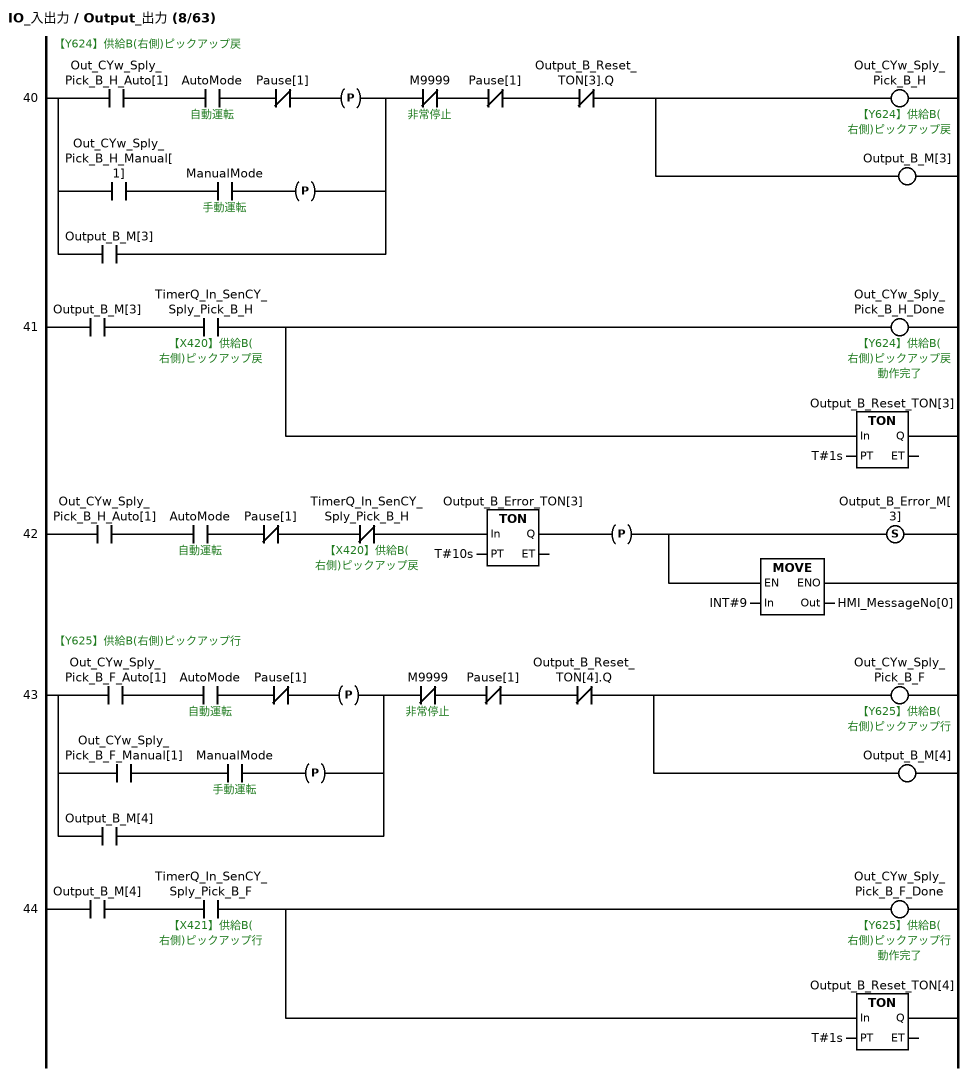
(* [picture p57: IO_入出力 / Output_出力, rungs 40-44] *)
(* Rung 40: 【Y624】供給B(右側)ピックアップ戻 *)
_e33(CLK := Out_CYw_Sply_Pick_B_H_Auto[1] AND AutoMode AND NOT Pause[1]);
_e34(CLK := Out_CYw_Sply_Pick_B_H_Manual[1] AND ManualMode);
_p35 := (_e33.Q OR _e34.Q OR Output_B_M[3]) AND NOT M9999 AND NOT Pause[1] AND NOT Output_B_Reset_TON[3].Q;
Out_CYw_Sply_Pick_B_H := _p35;
Output_B_M[3] := _p35;
(* Rung 41 *)
Out_CYw_Sply_Pick_B_H_Done := Output_B_M[3] AND TimerQ_In_SenCY_Sply_Pick_B_H;
Output_B_Reset_TON[3](In := Output_B_M[3] AND TimerQ_In_SenCY_Sply_Pick_B_H, PT := T#1s);
(* Rung 42 *)
Output_B_Error_TON[3](In := Out_CYw_Sply_Pick_B_H_Auto[1] AND AutoMode AND NOT Pause[1] AND NOT TimerQ_In_SenCY_Sply_Pick_B_H, PT := T#10s);
_e36(CLK := Output_B_Error_TON[3].Q);
IF _e36.Q THEN
    Output_B_Error_M[3] := TRUE;
    HMI_MessageNo[0] := INT#9;
END_IF;
(* Rung 43: 【Y625】供給B(右側)ピックアップ行 *)
_e37(CLK := Out_CYw_Sply_Pick_B_F_Auto[1] AND AutoMode AND NOT Pause[1]);
_e38(CLK := Out_CYw_Sply_Pick_B_F_Manual[1] AND ManualMode);
_p39 := (_e37.Q OR _e38.Q OR Output_B_M[4]) AND NOT M9999 AND NOT Pause[1] AND NOT Output_B_Reset_TON[4].Q;
Out_CYw_Sply_Pick_B_F := _p39;
Output_B_M[4] := _p39;
(* Rung 44 *)
Out_CYw_Sply_Pick_B_F_Done := Output_B_M[4] AND TimerQ_In_SenCY_Sply_Pick_B_F;
Output_B_Reset_TON[4](In := Output_B_M[4] AND TimerQ_In_SenCY_Sply_Pick_B_F, PT := T#1s);

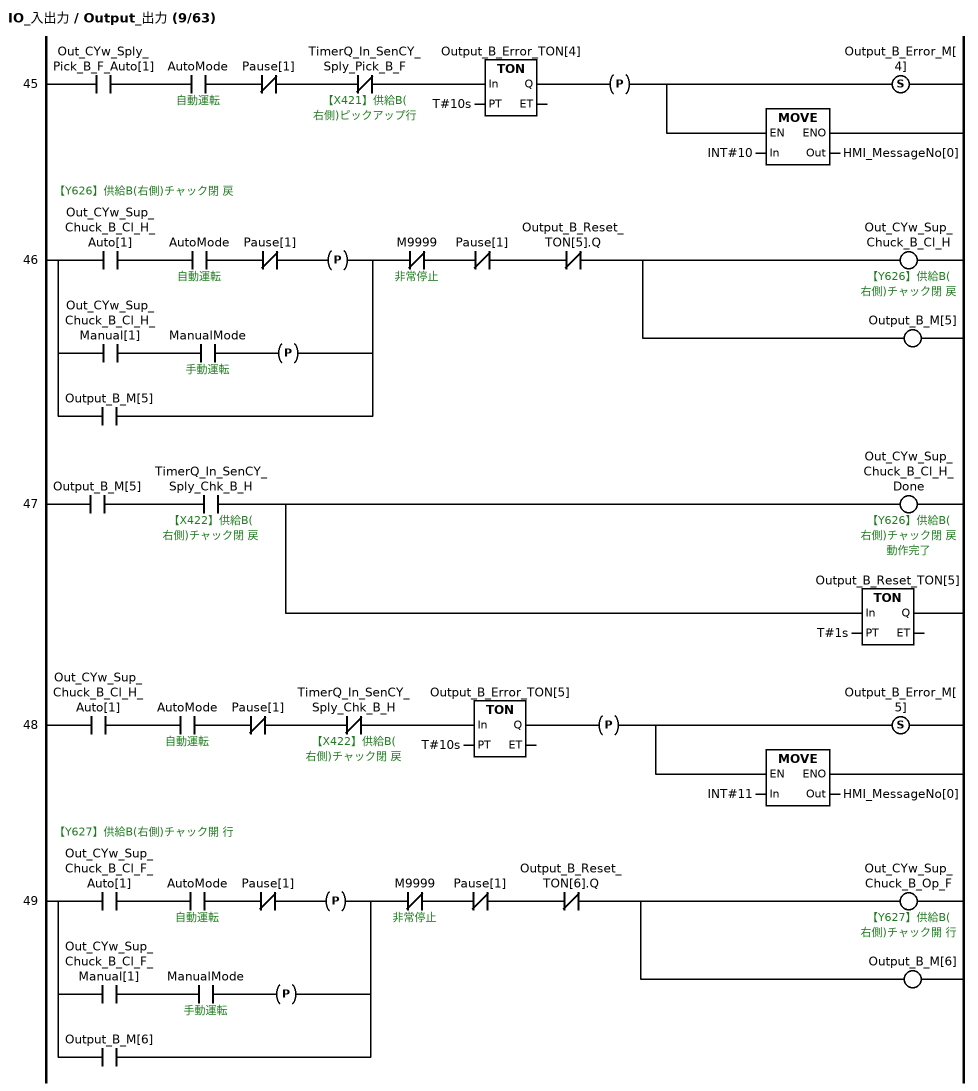
(* Rung 45 *)
Output_B_Error_TON[4](In := Out_CYw_Sply_Pick_B_F_Auto[1] AND AutoMode AND NOT Pause[1] AND NOT TimerQ_In_SenCY_Sply_Pick_B_F, PT := T#10s);
_e40(CLK := Output_B_Error_TON[4].Q);
IF _e40.Q THEN
    Output_B_Error_M[4] := TRUE;
    HMI_MessageNo[0] := INT#10;
END_IF;
(* Rung 46: 【Y626】供給B(右側)チャック閉 戻 *)
_e41(CLK := Out_CYw_Sup_Chuck_B_Cl_H_Auto[1] AND AutoMode AND NOT Pause[1]);
_e42(CLK := Out_CYw_Sup_Chuck_B_Cl_H_Manual[1] AND ManualMode);
_p43 := (_e41.Q OR _e42.Q OR Output_B_M[5]) AND NOT M9999 AND NOT Pause[1] AND NOT Output_B_Reset_TON[5].Q;
Out_CYw_Sup_Chuck_B_Cl_H := _p43;
Output_B_M[5] := _p43;
(* Rung 47 *)
Out_CYw_Sup_Chuck_B_Cl_H_Done := Output_B_M[5] AND TimerQ_In_SenCY_Sply_Chk_B_H;
Output_B_Reset_TON[5](In := Output_B_M[5] AND TimerQ_In_SenCY_Sply_Chk_B_H, PT := T#1s);
(* Rung 48 *)
Output_B_Error_TON[5](In := Out_CYw_Sup_Chuck_B_Cl_H_Auto[1] AND AutoMode AND NOT Pause[1] AND NOT TimerQ_In_SenCY_Sply_Chk_B_H, PT := T#10s);
_e44(CLK := Output_B_Error_TON[5].Q);
IF _e44.Q THEN
    Output_B_Error_M[5] := TRUE;
    HMI_MessageNo[0] := INT#11;
END_IF;
(* Rung 49: 【Y627】供給B(右側)チャック開 行 *)
_e45(CLK := Out_CYw_Sup_Chuck_B_Cl_F_Auto[1] AND AutoMode AND NOT Pause[1]);
_e46(CLK := Out_CYw_Sup_Chuck_B_Cl_F_Manual[1] AND ManualMode);
_p47 := (_e45.Q OR _e46.Q OR Output_B_M[6]) AND NOT M9999 AND NOT Pause[1] AND NOT Output_B_Reset_TON[6].Q;
Out_CYw_Sup_Chuck_B_Op_F := _p47;
Output_B_M[6] := _p47;

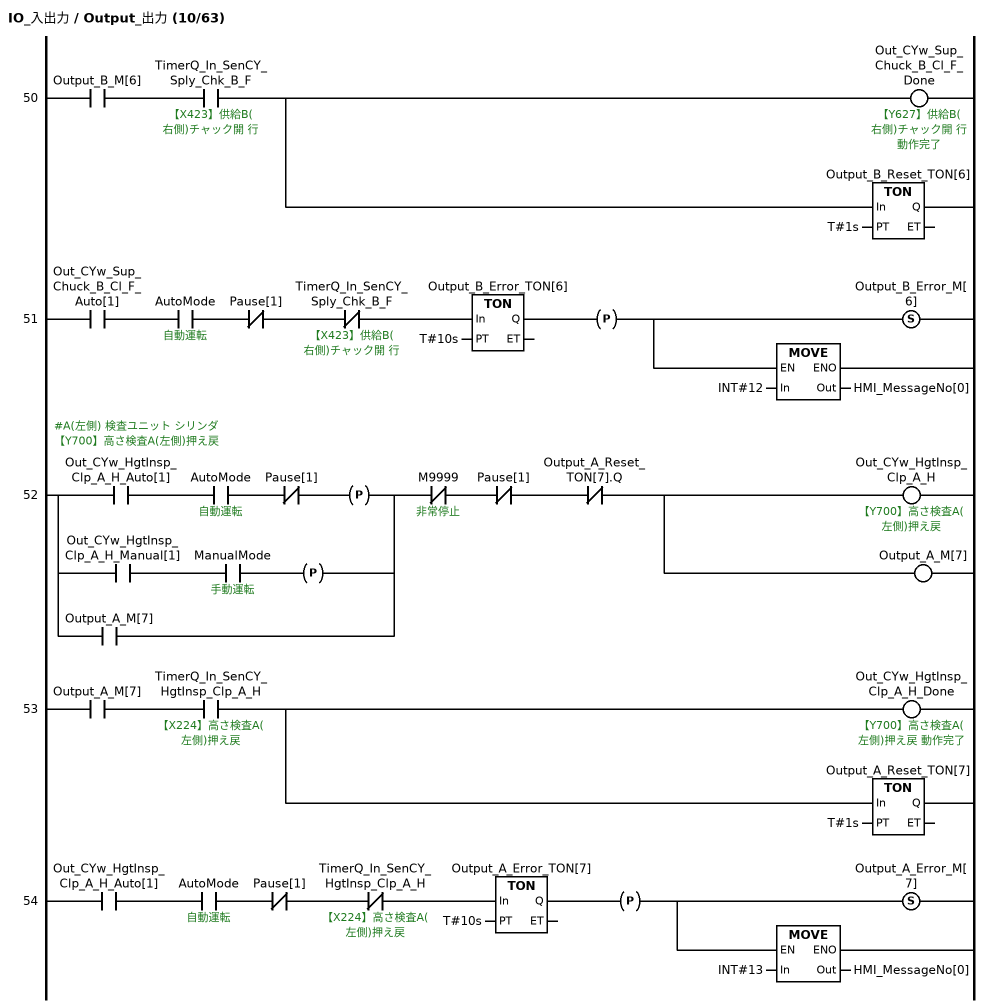
(* Rung 50 *)
Out_CYw_Sup_Chuck_B_Cl_F_Done := Output_B_M[6] AND TimerQ_In_SenCY_Sply_Chk_B_F;
Output_B_Reset_TON[6](In := Output_B_M[6] AND TimerQ_In_SenCY_Sply_Chk_B_F, PT := T#1s);
(* Rung 51 *)
Output_B_Error_TON[6](In := Out_CYw_Sup_Chuck_B_Cl_F_Auto[1] AND AutoMode AND NOT Pause[1] AND NOT TimerQ_In_SenCY_Sply_Chk_B_F, PT := T#10s);
_e48(CLK := Output_B_Error_TON[6].Q);
IF _e48.Q THEN
    Output_B_Error_M[6] := TRUE;
    HMI_MessageNo[0] := INT#12;
END_IF;
(* Rung 52: #A(左側) 検査ユニット シリンダ / 【Y700】高さ検査A(左側)押え戻 *)
_e49(CLK := Out_CYw_HgtInsp_Clp_A_H_Auto[1] AND AutoMode AND NOT Pause[1]);
_e50(CLK := Out_CYw_HgtInsp_Clp_A_H_Manual[1] AND ManualMode);
_p51 := (_e49.Q OR _e50.Q OR Output_A_M[7]) AND NOT M9999 AND NOT Pause[1] AND NOT Output_A_Reset_TON[7].Q;
Out_CYw_HgtInsp_Clp_A_H := _p51;
Output_A_M[7] := _p51;
(* Rung 53 *)
_p52 := Output_A_M[7] AND TimerQ_In_SenCY_HgtInsp_Clp_A_H;
Out_CYw_HgtInsp_Clp_A_H_Done := _p52;
Output_A_Reset_TON[7](In := _p52, PT := T#1s);
(* Rung 54 *)
Output_A_Error_TON[7](In := Out_CYw_HgtInsp_Clp_A_H_Auto[1] AND AutoMode AND NOT Pause[1] AND NOT TimerQ_In_SenCY_HgtInsp_Clp_A_H, PT := T#10s);
_e53(CLK := Output_A_Error_TON[7].Q);
IF _e53.Q THEN
    Output_A_Error_M[7] := TRUE;
    HMI_MessageNo[0] := INT#13;
END_IF;

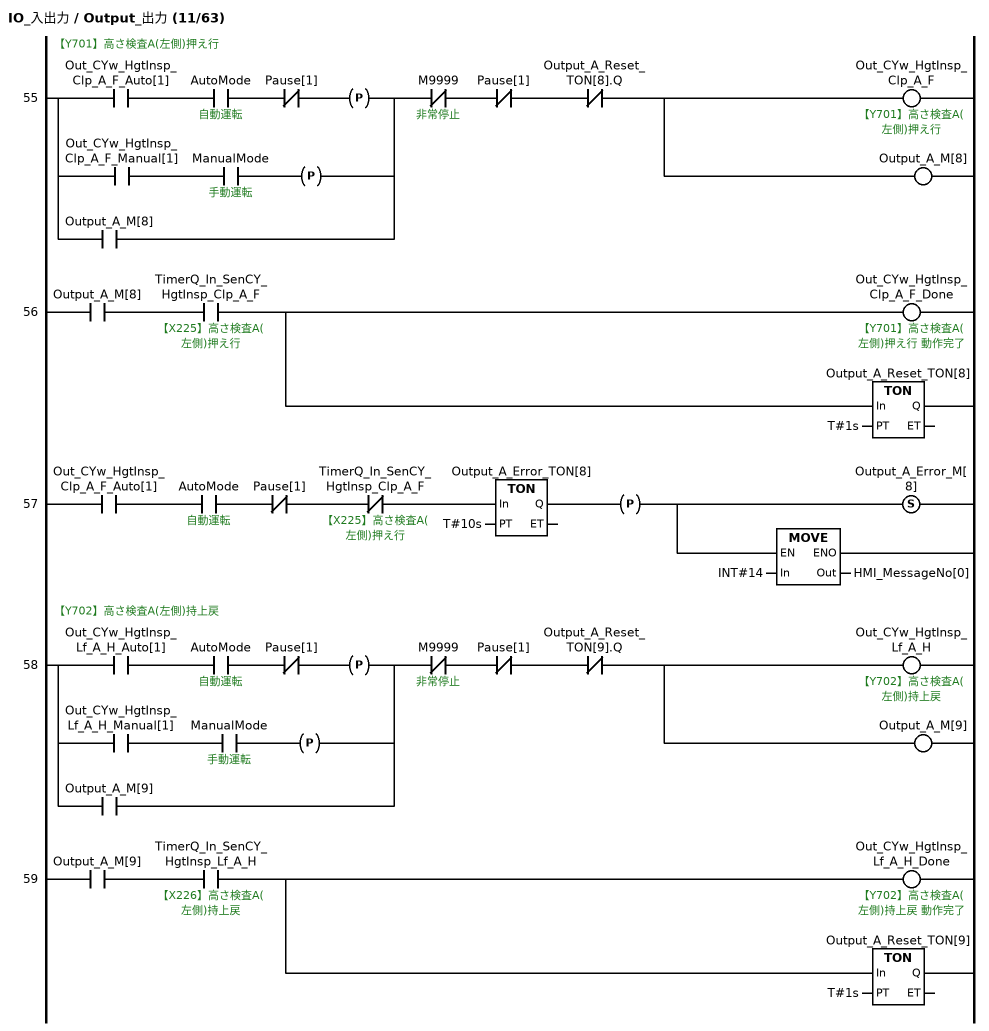
(* Rung 55: 【Y701】高さ検査A(左側)押え行 *)
_e54(CLK := Out_CYw_HgtInsp_Clp_A_F_Auto[1] AND AutoMode AND NOT Pause[1]);
_e55(CLK := Out_CYw_HgtInsp_Clp_A_F_Manual[1] AND ManualMode);
_p56 := (_e54.Q OR _e55.Q OR Output_A_M[8]) AND NOT M9999 AND NOT Pause[1] AND NOT Output_A_Reset_TON[8].Q;
Out_CYw_HgtInsp_Clp_A_F := _p56;
Output_A_M[8] := _p56;
(* Rung 56 *)
_p57 := Output_A_M[8] AND TimerQ_In_SenCY_HgtInsp_Clp_A_F;
Out_CYw_HgtInsp_Clp_A_F_Done := _p57;
Output_A_Reset_TON[8](In := _p57, PT := T#1s);
(* Rung 57 *)
Output_A_Error_TON[8](In := Out_CYw_HgtInsp_Clp_A_F_Auto[1] AND AutoMode AND NOT Pause[1] AND NOT TimerQ_In_SenCY_HgtInsp_Clp_A_F, PT := T#10s);
_e58(CLK := Output_A_Error_TON[8].Q);
IF _e58.Q THEN
    Output_A_Error_M[8] := TRUE;
    HMI_MessageNo[0] := INT#14;
END_IF;
(* Rung 58: 【Y702】高さ検査A(左側)持上戻 *)
_e59(CLK := Out_CYw_HgtInsp_Lf_A_H_Auto[1] AND AutoMode AND NOT Pause[1]);
_e60(CLK := Out_CYw_HgtInsp_Lf_A_H_Manual[1] AND ManualMode);
_p61 := (_e59.Q OR _e60.Q OR Output_A_M[9]) AND NOT M9999 AND NOT Pause[1] AND NOT Output_A_Reset_TON[9].Q;
Out_CYw_HgtInsp_Lf_A_H := _p61;
Output_A_M[9] := _p61;
(* Rung 59 *)
Out_CYw_HgtInsp_Lf_A_H_Done := Output_A_M[9] AND TimerQ_In_SenCY_HgtInsp_Lf_A_H;
Output_A_Reset_TON[9](In := Output_A_M[9] AND TimerQ_In_SenCY_HgtInsp_Lf_A_H, PT := T#1s);

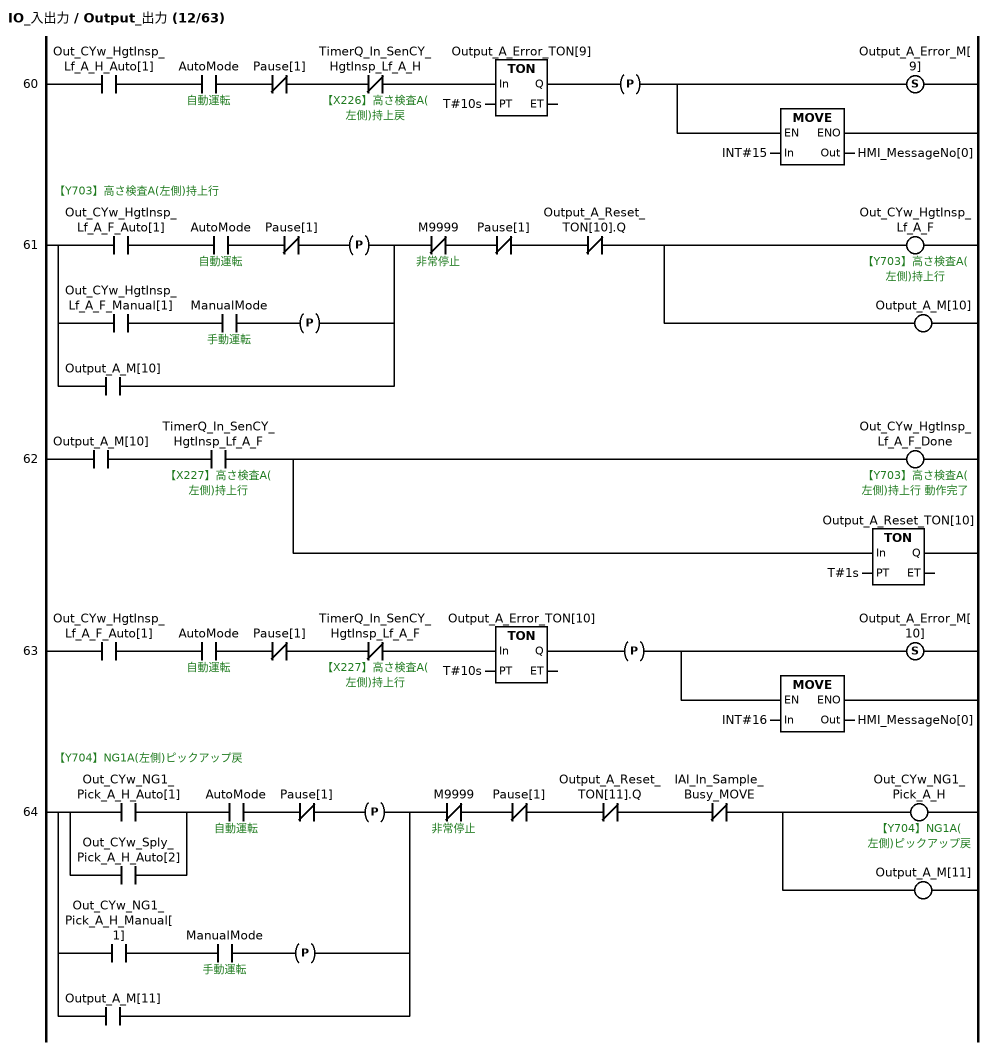
(* Rung 60 *)
Output_A_Error_TON[9](In := Out_CYw_HgtInsp_Lf_A_H_Auto[1] AND AutoMode AND NOT Pause[1] AND NOT TimerQ_In_SenCY_HgtInsp_Lf_A_H, PT := T#10s);
_e62(CLK := Output_A_Error_TON[9].Q);
IF _e62.Q THEN
    Output_A_Error_M[9] := TRUE;
    HMI_MessageNo[0] := INT#15;
END_IF;
(* Rung 61: 【Y703】高さ検査A(左側)持上行 *)
_e63(CLK := Out_CYw_HgtInsp_Lf_A_F_Auto[1] AND AutoMode AND NOT Pause[1]);
_e64(CLK := Out_CYw_HgtInsp_Lf_A_F_Manual[1] AND ManualMode);
_p65 := (_e63.Q OR _e64.Q OR Output_A_M[10]) AND NOT M9999 AND NOT Pause[1] AND NOT Output_A_Reset_TON[10].Q;
Out_CYw_HgtInsp_Lf_A_F := _p65;
Output_A_M[10] := _p65;
(* Rung 62 *)
_p66 := Output_A_M[10] AND TimerQ_In_SenCY_HgtInsp_Lf_A_F;
Out_CYw_HgtInsp_Lf_A_F_Done := _p66;
Output_A_Reset_TON[10](In := _p66, PT := T#1s);
(* Rung 63 *)
Output_A_Error_TON[10](In := Out_CYw_HgtInsp_Lf_A_F_Auto[1] AND AutoMode AND NOT Pause[1] AND NOT TimerQ_In_SenCY_HgtInsp_Lf_A_F, PT := T#10s);
_e67(CLK := Output_A_Error_TON[10].Q);
IF _e67.Q THEN
    Output_A_Error_M[10] := TRUE;
    HMI_MessageNo[0] := INT#16;
END_IF;
(* Rung 64: 【Y704】NG1A(左側)ピックアップ戻 *)
_e68(CLK := (Out_CYw_NG1_Pick_A_H_Auto[1] OR Out_CYw_Sply_Pick_A_H_Auto[2]) AND AutoMode AND NOT Pause[1]);
_e69(CLK := Out_CYw_NG1_Pick_A_H_Manual[1] AND ManualMode);
_p70 := (_e68.Q OR _e69.Q OR Output_A_M[11]) AND NOT M9999 AND NOT Pause[1] AND NOT Output_A_Reset_TON[11].Q AND NOT IAI_In_Sample_Busy_MOVE;
Out_CYw_NG1_Pick_A_H := _p70;
Output_A_M[11] := _p70;

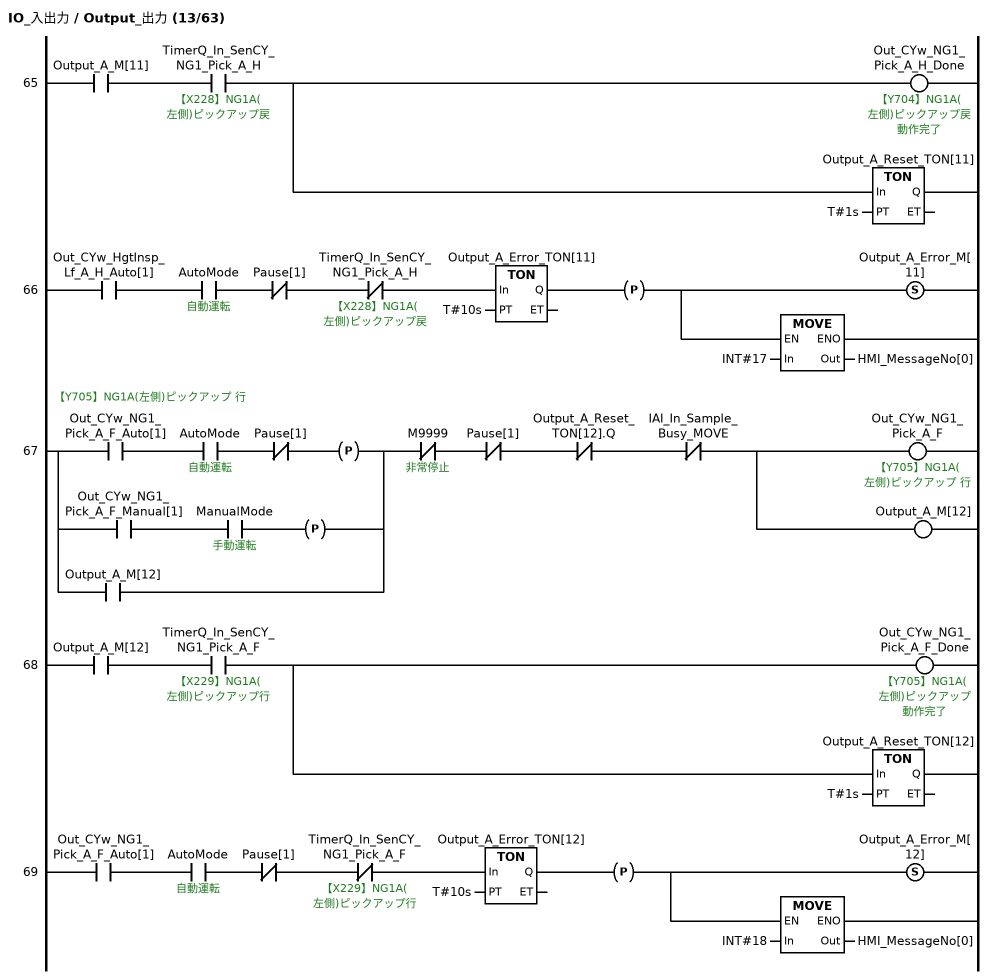
(* Rung 65 *)
Out_CYw_NG1_Pick_A_H_Done := Output_A_M[11] AND TimerQ_In_SenCY_NG1_Pick_A_H;
Output_A_Reset_TON[11](In := Output_A_M[11] AND TimerQ_In_SenCY_NG1_Pick_A_H, PT := T#1s);
(* Rung 66 *)
Output_A_Error_TON[11](In := Out_CYw_HgtInsp_Lf_A_H_Auto[1] AND AutoMode AND NOT Pause[1] AND NOT TimerQ_In_SenCY_NG1_Pick_A_H, PT := T#10s);
_e71(CLK := Output_A_Error_TON[11].Q);
IF _e71.Q THEN
    Output_A_Error_M[11] := TRUE;
    HMI_MessageNo[0] := INT#17;
END_IF;
(* Rung 67: 【Y705】NG1A(左側)ピックアップ 行 *)
_e72(CLK := Out_CYw_NG1_Pick_A_F_Auto[1] AND AutoMode AND NOT Pause[1]);
_e73(CLK := Out_CYw_NG1_Pick_A_F_Manual[1] AND ManualMode);
_p74 := (_e72.Q OR _e73.Q OR Output_A_M[12]) AND NOT M9999 AND NOT Pause[1] AND NOT Output_A_Reset_TON[12].Q AND NOT IAI_In_Sample_Busy_MOVE;
Out_CYw_NG1_Pick_A_F := _p74;
Output_A_M[12] := _p74;
(* Rung 68 *)
Out_CYw_NG1_Pick_A_F_Done := Output_A_M[12] AND TimerQ_In_SenCY_NG1_Pick_A_F;
Output_A_Reset_TON[12](In := Output_A_M[12] AND TimerQ_In_SenCY_NG1_Pick_A_F, PT := T#1s);
(* Rung 69 *)
Output_A_Error_TON[12](In := Out_CYw_NG1_Pick_A_F_Auto[1] AND AutoMode AND NOT Pause[1] AND NOT TimerQ_In_SenCY_NG1_Pick_A_F, PT := T#10s);
_e75(CLK := Output_A_Error_TON[12].Q);
IF _e75.Q THEN
    Output_A_Error_M[12] := TRUE;
    HMI_MessageNo[0] := INT#18;
END_IF;

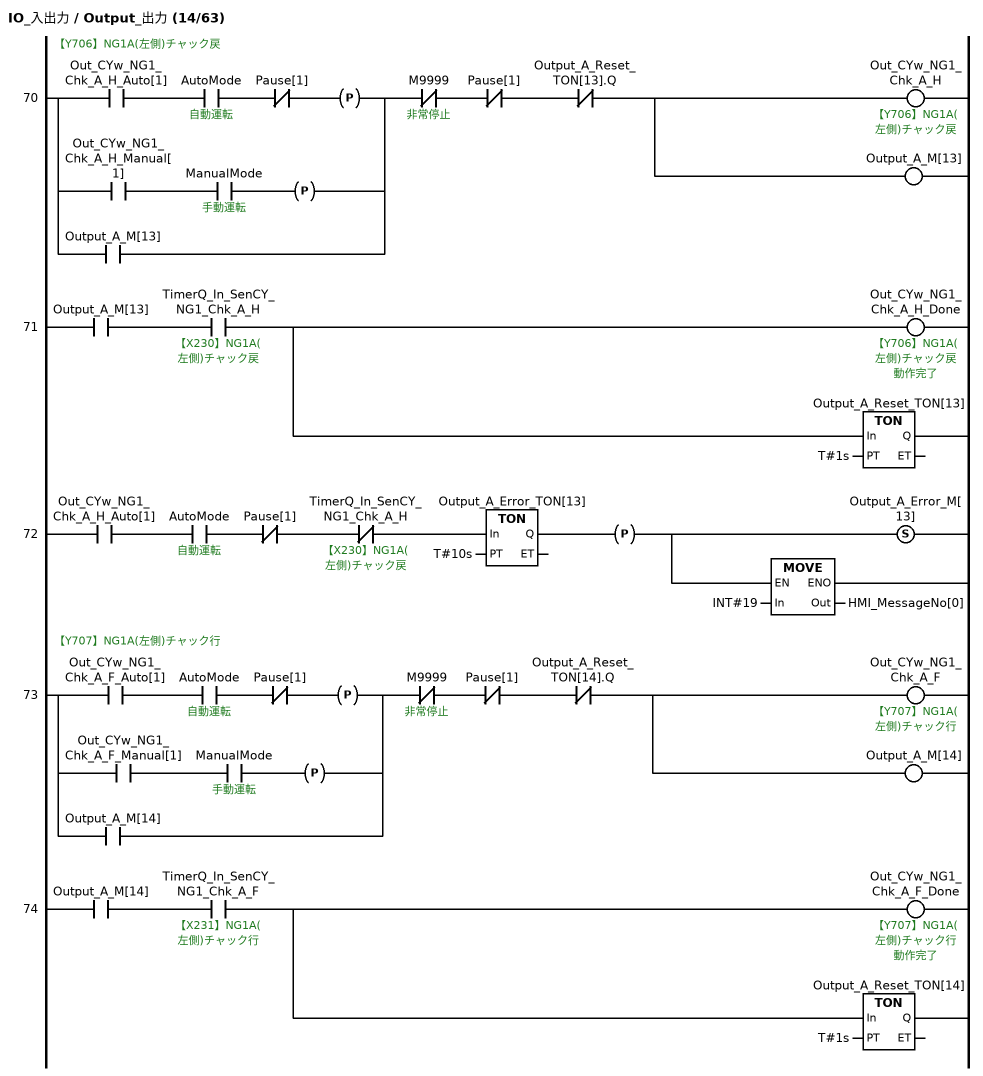
(* Rung 70: 【Y706】NG1A(左側)チャック戻 *)
_e76(CLK := Out_CYw_NG1_Chk_A_H_Auto[1] AND AutoMode AND NOT Pause[1]);
_e77(CLK := Out_CYw_NG1_Chk_A_H_Manual[1] AND ManualMode);
_p78 := (_e76.Q OR _e77.Q OR Output_A_M[13]) AND NOT M9999 AND NOT Pause[1] AND NOT Output_A_Reset_TON[13].Q;
Out_CYw_NG1_Chk_A_H := _p78;
Output_A_M[13] := _p78;
(* Rung 71 *)
Out_CYw_NG1_Chk_A_H_Done := Output_A_M[13] AND TimerQ_In_SenCY_NG1_Chk_A_H;
Output_A_Reset_TON[13](In := Output_A_M[13] AND TimerQ_In_SenCY_NG1_Chk_A_H, PT := T#1s);
(* Rung 72 *)
Output_A_Error_TON[13](In := Out_CYw_NG1_Chk_A_H_Auto[1] AND AutoMode AND NOT Pause[1] AND NOT TimerQ_In_SenCY_NG1_Chk_A_H, PT := T#10s);
_e79(CLK := Output_A_Error_TON[13].Q);
IF _e79.Q THEN
    Output_A_Error_M[13] := TRUE;
    HMI_MessageNo[0] := INT#19;
END_IF;
(* Rung 73: 【Y707】NG1A(左側)チャック行 *)
_e80(CLK := Out_CYw_NG1_Chk_A_F_Auto[1] AND AutoMode AND NOT Pause[1]);
_e81(CLK := Out_CYw_NG1_Chk_A_F_Manual[1] AND ManualMode);
_p82 := (_e80.Q OR _e81.Q OR Output_A_M[14]) AND NOT M9999 AND NOT Pause[1] AND NOT Output_A_Reset_TON[14].Q;
Out_CYw_NG1_Chk_A_F := _p82;
Output_A_M[14] := _p82;
(* Rung 74 *)
Out_CYw_NG1_Chk_A_F_Done := Output_A_M[14] AND TimerQ_In_SenCY_NG1_Chk_A_F;
Output_A_Reset_TON[14](In := Output_A_M[14] AND TimerQ_In_SenCY_NG1_Chk_A_F, PT := T#1s);

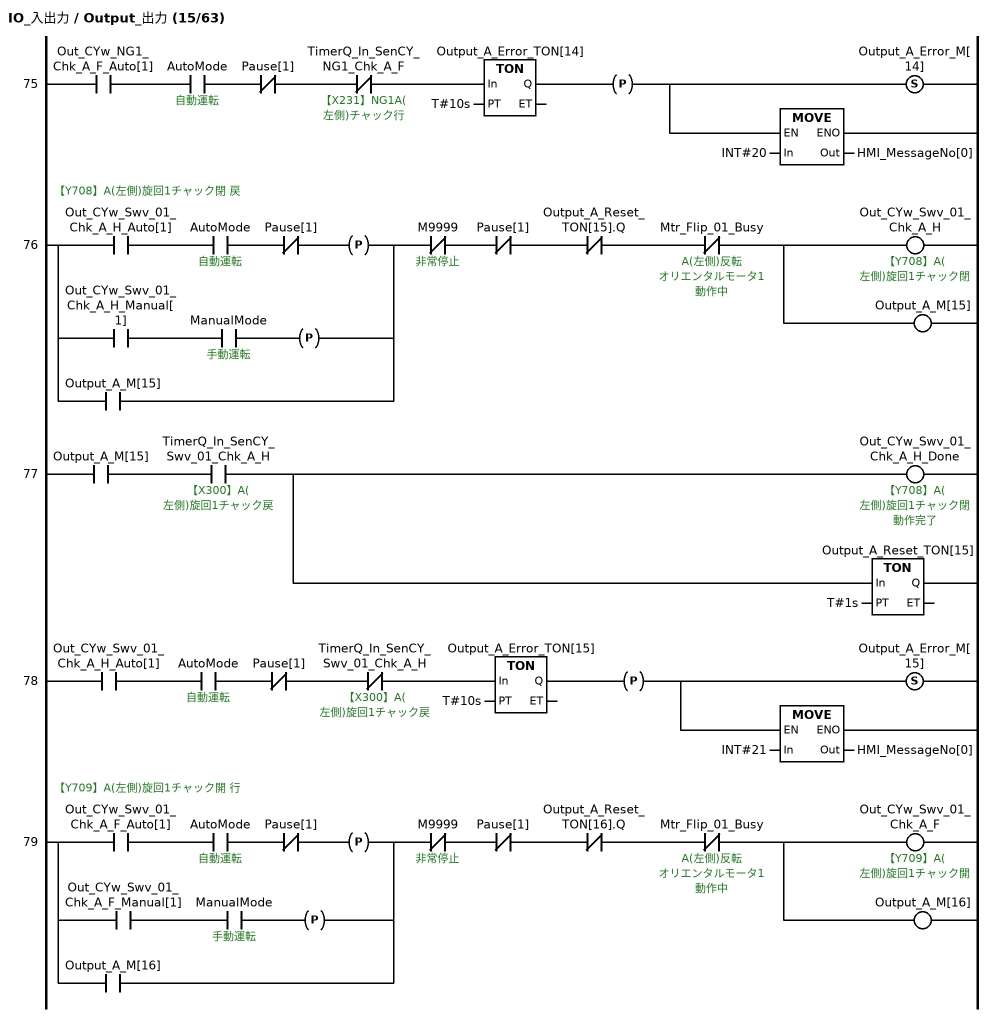
(* Rung 75 *)
Output_A_Error_TON[14](In := Out_CYw_NG1_Chk_A_F_Auto[1] AND AutoMode AND NOT Pause[1] AND NOT TimerQ_In_SenCY_NG1_Chk_A_F, PT := T#10s);
_e83(CLK := Output_A_Error_TON[14].Q);
IF _e83.Q THEN
    Output_A_Error_M[14] := TRUE;
    HMI_MessageNo[0] := INT#20;
END_IF;
(* Rung 76: 【Y708】A(左側)旋回1チャック閉 戻 *)
_e84(CLK := Out_CYw_Swv_01_Chk_A_H_Auto[1] AND AutoMode AND NOT Pause[1]);
_e85(CLK := Out_CYw_Swv_01_Chk_A_H_Manual[1] AND ManualMode);
_p86 := (_e84.Q OR _e85.Q OR Output_A_M[15]) AND NOT M9999 AND NOT Pause[1] AND NOT Output_A_Reset_TON[15].Q AND NOT Mtr_Flip_01_Busy;
Out_CYw_Swv_01_Chk_A_H := _p86;
Output_A_M[15] := _p86;
(* Rung 77 *)
_p87 := Output_A_M[15] AND TimerQ_In_SenCY_Swv_01_Chk_A_H;
Out_CYw_Swv_01_Chk_A_H_Done := _p87;
Output_A_Reset_TON[15](In := _p87, PT := T#1s);
(* Rung 78 *)
Output_A_Error_TON[15](In := Out_CYw_Swv_01_Chk_A_H_Auto[1] AND AutoMode AND NOT Pause[1] AND NOT TimerQ_In_SenCY_Swv_01_Chk_A_H, PT := T#10s);
_e88(CLK := Output_A_Error_TON[15].Q);
IF _e88.Q THEN
    Output_A_Error_M[15] := TRUE;
    HMI_MessageNo[0] := INT#21;
END_IF;
(* Rung 79: 【Y709】A(左側)旋回1チャック開 行 *)
_e89(CLK := Out_CYw_Swv_01_Chk_A_F_Auto[1] AND AutoMode AND NOT Pause[1]);
_e90(CLK := Out_CYw_Swv_01_Chk_A_F_Manual[1] AND ManualMode);
_p91 := (_e89.Q OR _e90.Q OR Output_A_M[16]) AND NOT M9999 AND NOT Pause[1] AND NOT Output_A_Reset_TON[16].Q AND NOT Mtr_Flip_01_Busy;
Out_CYw_Swv_01_Chk_A_F := _p91;
Output_A_M[16] := _p91;

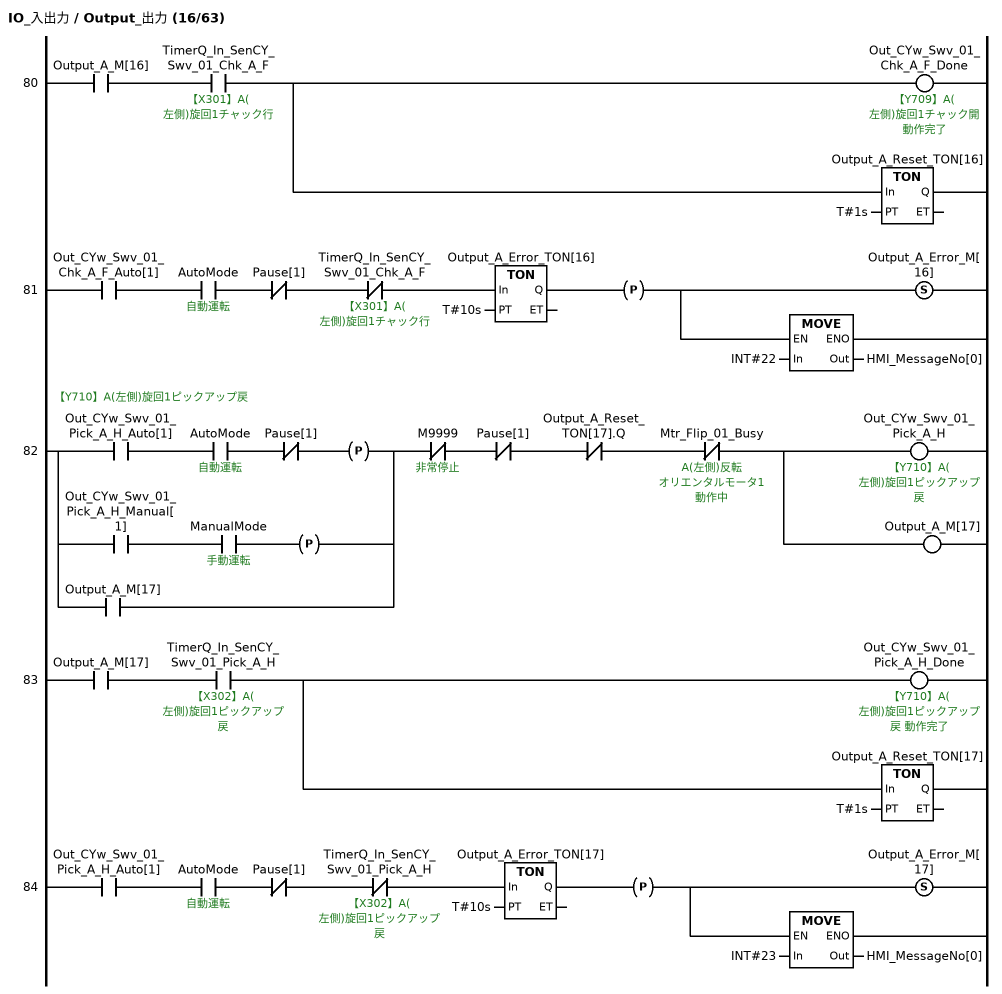
(* Rung 80 *)
_p92 := Output_A_M[16] AND TimerQ_In_SenCY_Swv_01_Chk_A_F;
Out_CYw_Swv_01_Chk_A_F_Done := _p92;
Output_A_Reset_TON[16](In := _p92, PT := T#1s);
(* Rung 81 *)
Output_A_Error_TON[16](In := Out_CYw_Swv_01_Chk_A_F_Auto[1] AND AutoMode AND NOT Pause[1] AND NOT TimerQ_In_SenCY_Swv_01_Chk_A_F, PT := T#10s);
_e93(CLK := Output_A_Error_TON[16].Q);
IF _e93.Q THEN
    Output_A_Error_M[16] := TRUE;
    HMI_MessageNo[0] := INT#22;
END_IF;
(* Rung 82: 【Y710】A(左側)旋回1ピックアップ戻 *)
_e94(CLK := Out_CYw_Swv_01_Pick_A_H_Auto[1] AND AutoMode AND NOT Pause[1]);
_e95(CLK := Out_CYw_Swv_01_Pick_A_H_Manual[1] AND ManualMode);
_p96 := (_e94.Q OR _e95.Q OR Output_A_M[17]) AND NOT M9999 AND NOT Pause[1] AND NOT Output_A_Reset_TON[17].Q AND NOT Mtr_Flip_01_Busy;
Out_CYw_Swv_01_Pick_A_H := _p96;
Output_A_M[17] := _p96;
(* Rung 83 *)
_p97 := Output_A_M[17] AND TimerQ_In_SenCY_Swv_01_Pick_A_H;
Out_CYw_Swv_01_Pick_A_H_Done := _p97;
Output_A_Reset_TON[17](In := _p97, PT := T#1s);
(* Rung 84 *)
Output_A_Error_TON[17](In := Out_CYw_Swv_01_Pick_A_H_Auto[1] AND AutoMode AND NOT Pause[1] AND NOT TimerQ_In_SenCY_Swv_01_Pick_A_H, PT := T#10s);
_e98(CLK := Output_A_Error_TON[17].Q);
IF _e98.Q THEN
    Output_A_Error_M[17] := TRUE;
    HMI_MessageNo[0] := INT#23;
END_IF;

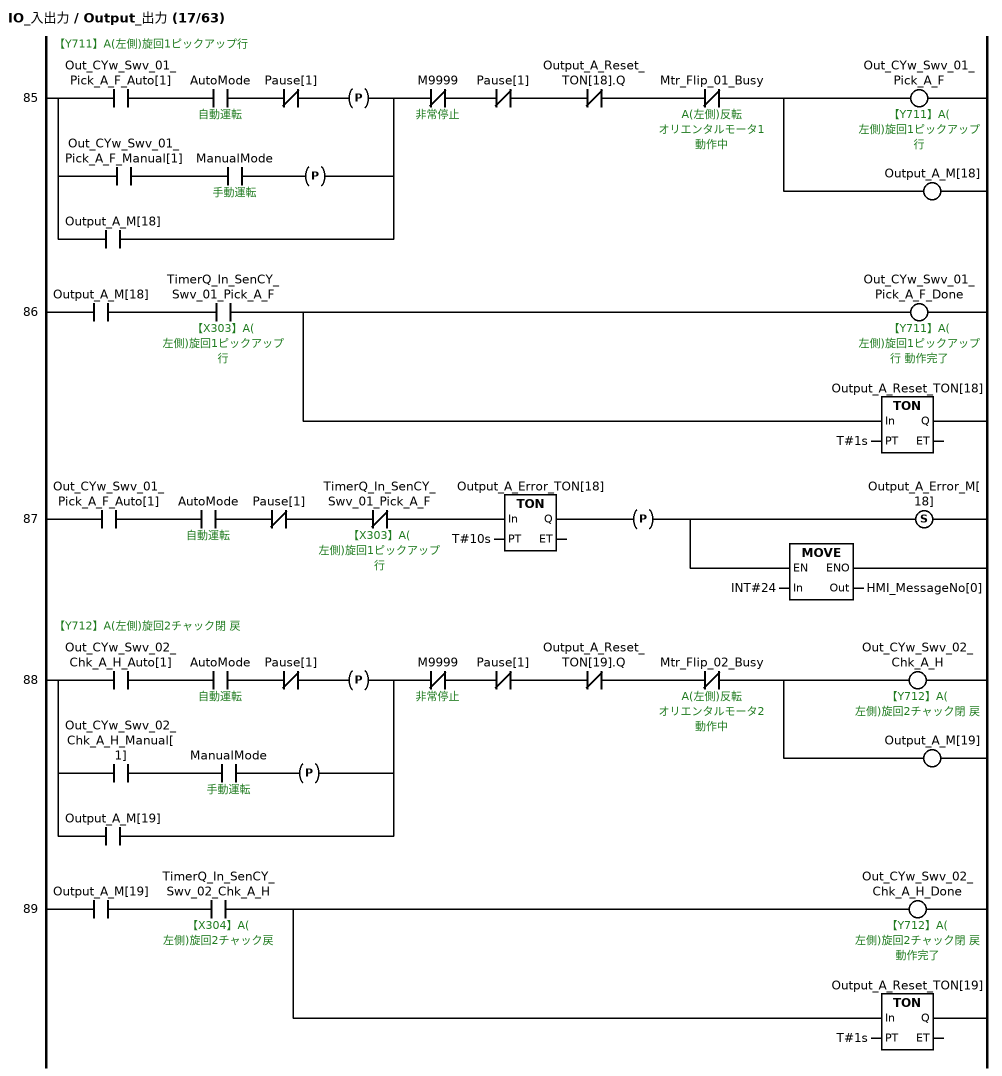
(* Rung 85: 【Y711】A(左側)旋回1ピックアップ行 *)
_e99(CLK := Out_CYw_Swv_01_Pick_A_F_Auto[1] AND AutoMode AND NOT Pause[1]);
_e100(CLK := Out_CYw_Swv_01_Pick_A_F_Manual[1] AND ManualMode);
_p101 := (_e99.Q OR _e100.Q OR Output_A_M[18]) AND NOT M9999 AND NOT Pause[1] AND NOT Output_A_Reset_TON[18].Q AND NOT Mtr_Flip_01_Busy;
Out_CYw_Swv_01_Pick_A_F := _p101;
Output_A_M[18] := _p101;
(* Rung 86 *)
_p102 := Output_A_M[18] AND TimerQ_In_SenCY_Swv_01_Pick_A_F;
Out_CYw_Swv_01_Pick_A_F_Done := _p102;
Output_A_Reset_TON[18](In := _p102, PT := T#1s);
(* Rung 87 *)
Output_A_Error_TON[18](In := Out_CYw_Swv_01_Pick_A_F_Auto[1] AND AutoMode AND NOT Pause[1] AND NOT TimerQ_In_SenCY_Swv_01_Pick_A_F, PT := T#10s);
_e103(CLK := Output_A_Error_TON[18].Q);
IF _e103.Q THEN
    Output_A_Error_M[18] := TRUE;
    HMI_MessageNo[0] := INT#24;
END_IF;
(* Rung 88: 【Y712】A(左側)旋回2チャック閉 戻 *)
_e104(CLK := Out_CYw_Swv_02_Chk_A_H_Auto[1] AND AutoMode AND NOT Pause[1]);
_e105(CLK := Out_CYw_Swv_02_Chk_A_H_Manual[1] AND ManualMode);
_p106 := (_e104.Q OR _e105.Q OR Output_A_M[19]) AND NOT M9999 AND NOT Pause[1] AND NOT Output_A_Reset_TON[19].Q AND NOT Mtr_Flip_02_Busy;
Out_CYw_Swv_02_Chk_A_H := _p106;
Output_A_M[19] := _p106;
(* Rung 89 *)
_p107 := Output_A_M[19] AND TimerQ_In_SenCY_Swv_02_Chk_A_H;
Out_CYw_Swv_02_Chk_A_H_Done := _p107;
Output_A_Reset_TON[19](In := _p107, PT := T#1s);

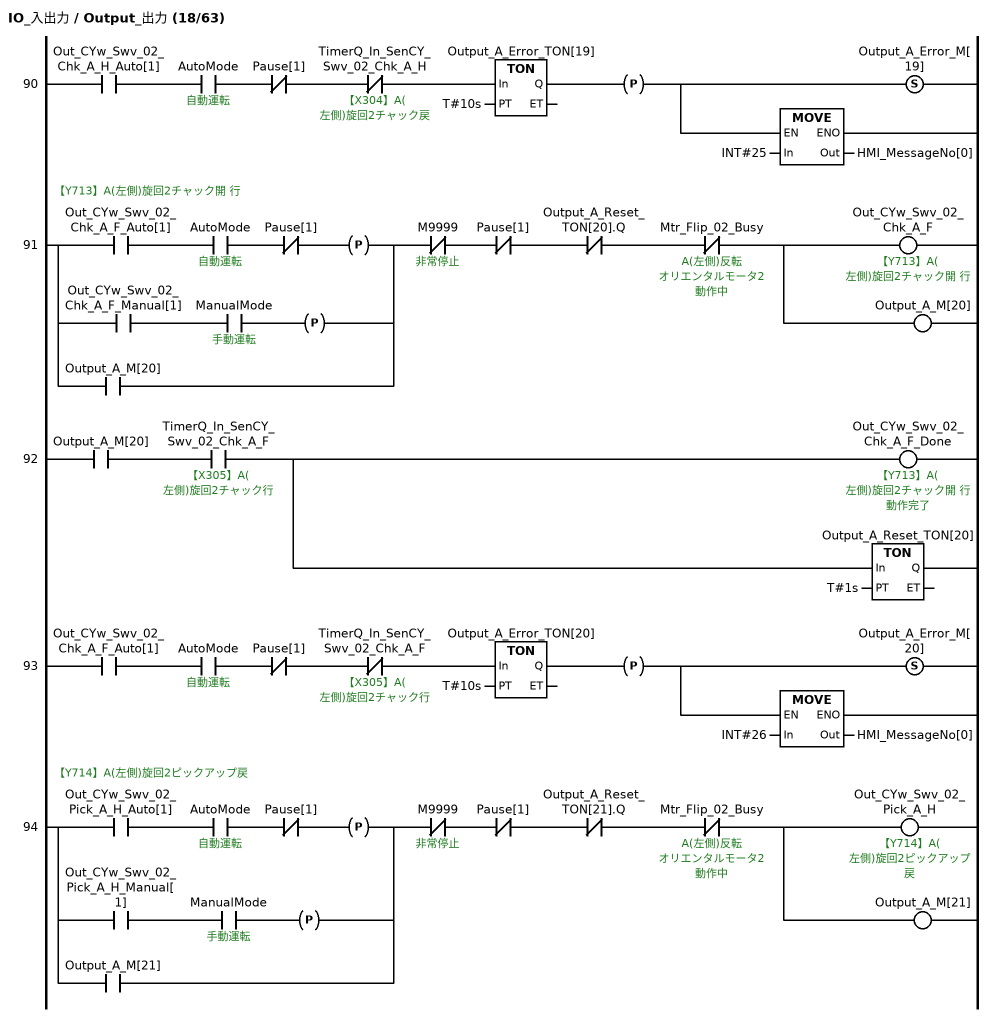
(* Rung 90 *)
Output_A_Error_TON[19](In := Out_CYw_Swv_02_Chk_A_H_Auto[1] AND AutoMode AND NOT Pause[1] AND NOT TimerQ_In_SenCY_Swv_02_Chk_A_H, PT := T#10s);
_e108(CLK := Output_A_Error_TON[19].Q);
IF _e108.Q THEN
    Output_A_Error_M[19] := TRUE;
    HMI_MessageNo[0] := INT#25;
END_IF;
(* Rung 91: 【Y713】A(左側)旋回2チャック開 行 *)
_e109(CLK := Out_CYw_Swv_02_Chk_A_F_Auto[1] AND AutoMode AND NOT Pause[1]);
_e110(CLK := Out_CYw_Swv_02_Chk_A_F_Manual[1] AND ManualMode);
_p111 := (_e109.Q OR _e110.Q OR Output_A_M[20]) AND NOT M9999 AND NOT Pause[1] AND NOT Output_A_Reset_TON[20].Q AND NOT Mtr_Flip_02_Busy;
Out_CYw_Swv_02_Chk_A_F := _p111;
Output_A_M[20] := _p111;
(* Rung 92 *)
_p112 := Output_A_M[20] AND TimerQ_In_SenCY_Swv_02_Chk_A_F;
Out_CYw_Swv_02_Chk_A_F_Done := _p112;
Output_A_Reset_TON[20](In := _p112, PT := T#1s);
(* Rung 93 *)
Output_A_Error_TON[20](In := Out_CYw_Swv_02_Chk_A_F_Auto[1] AND AutoMode AND NOT Pause[1] AND NOT TimerQ_In_SenCY_Swv_02_Chk_A_F, PT := T#10s);
_e113(CLK := Output_A_Error_TON[20].Q);
IF _e113.Q THEN
    Output_A_Error_M[20] := TRUE;
    HMI_MessageNo[0] := INT#26;
END_IF;
(* Rung 94: 【Y714】A(左側)旋回2ピックアップ戻 *)
_e114(CLK := Out_CYw_Swv_02_Pick_A_H_Auto[1] AND AutoMode AND NOT Pause[1]);
_e115(CLK := Out_CYw_Swv_02_Pick_A_H_Manual[1] AND ManualMode);
_p116 := (_e114.Q OR _e115.Q OR Output_A_M[21]) AND NOT M9999 AND NOT Pause[1] AND NOT Output_A_Reset_TON[21].Q AND NOT Mtr_Flip_02_Busy;
Out_CYw_Swv_02_Pick_A_H := _p116;
Output_A_M[21] := _p116;

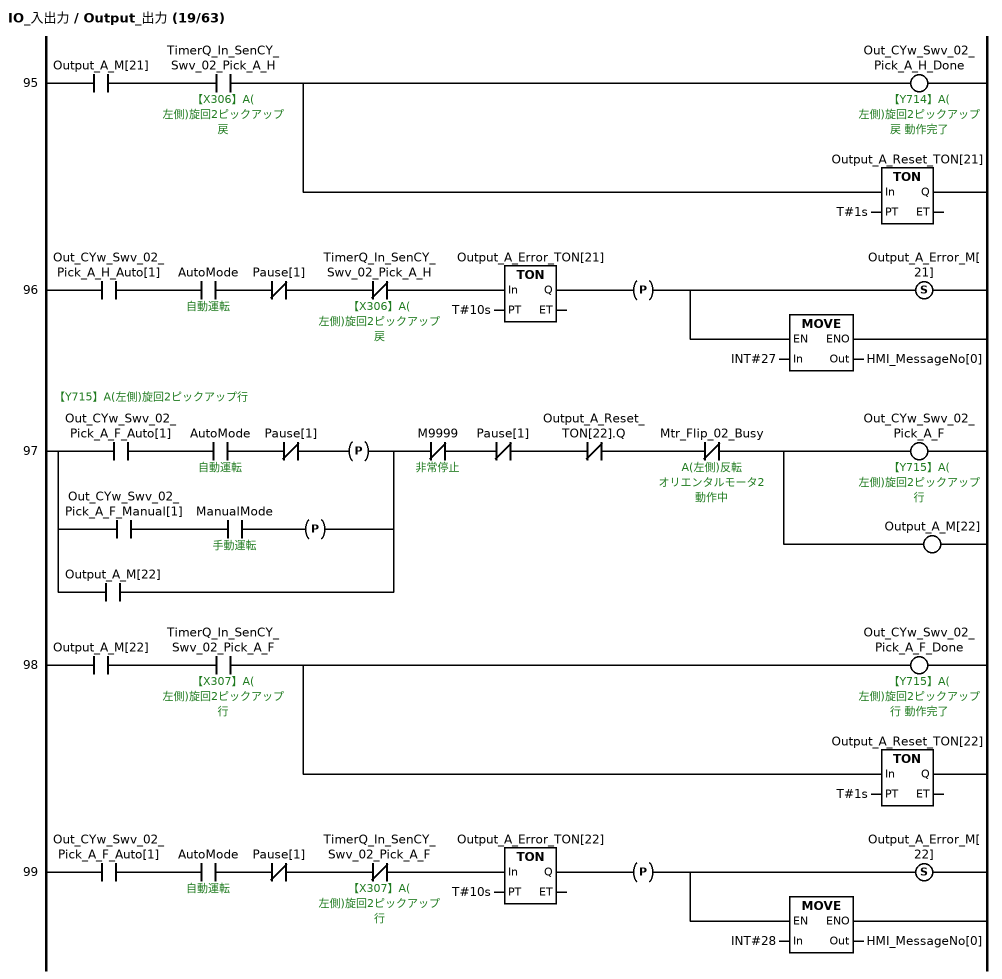
(* Rung 95 *)
_p117 := Output_A_M[21] AND TimerQ_In_SenCY_Swv_02_Pick_A_H;
Out_CYw_Swv_02_Pick_A_H_Done := _p117;
Output_A_Reset_TON[21](In := _p117, PT := T#1s);
(* Rung 96 *)
Output_A_Error_TON[21](In := Out_CYw_Swv_02_Pick_A_H_Auto[1] AND AutoMode AND NOT Pause[1] AND NOT TimerQ_In_SenCY_Swv_02_Pick_A_H, PT := T#10s);
_e118(CLK := Output_A_Error_TON[21].Q);
IF _e118.Q THEN
    Output_A_Error_M[21] := TRUE;
    HMI_MessageNo[0] := INT#27;
END_IF;
(* Rung 97: 【Y715】A(左側)旋回2ピックアップ行 *)
_e119(CLK := Out_CYw_Swv_02_Pick_A_F_Auto[1] AND AutoMode AND NOT Pause[1]);
_e120(CLK := Out_CYw_Swv_02_Pick_A_F_Manual[1] AND ManualMode);
_p121 := (_e119.Q OR _e120.Q OR Output_A_M[22]) AND NOT M9999 AND NOT Pause[1] AND NOT Output_A_Reset_TON[22].Q AND NOT Mtr_Flip_02_Busy;
Out_CYw_Swv_02_Pick_A_F := _p121;
Output_A_M[22] := _p121;
(* Rung 98 *)
_p122 := Output_A_M[22] AND TimerQ_In_SenCY_Swv_02_Pick_A_F;
Out_CYw_Swv_02_Pick_A_F_Done := _p122;
Output_A_Reset_TON[22](In := _p122, PT := T#1s);
(* Rung 99 *)
Output_A_Error_TON[22](In := Out_CYw_Swv_02_Pick_A_F_Auto[1] AND AutoMode AND NOT Pause[1] AND NOT TimerQ_In_SenCY_Swv_02_Pick_A_F, PT := T#10s);
_e123(CLK := Output_A_Error_TON[22].Q);
IF _e123.Q THEN
    Output_A_Error_M[22] := TRUE;
    HMI_MessageNo[0] := INT#28;
END_IF;

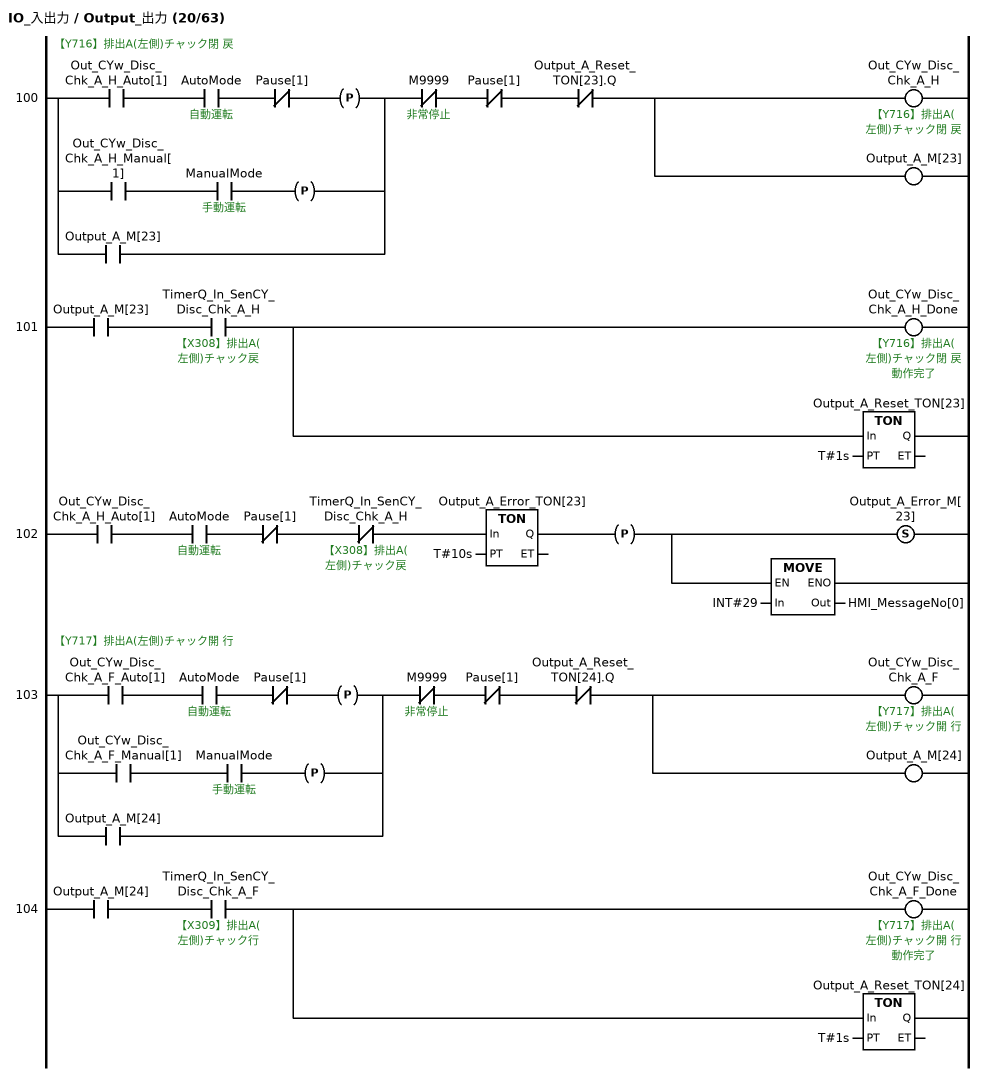
(* Rung 100: 【Y716】排出A(左側)チャック閉 戻 *)
_e124(CLK := Out_CYw_Disc_Chk_A_H_Auto[1] AND AutoMode AND NOT Pause[1]);
_e125(CLK := Out_CYw_Disc_Chk_A_H_Manual[1] AND ManualMode);
_p126 := (_e124.Q OR _e125.Q OR Output_A_M[23]) AND NOT M9999 AND NOT Pause[1] AND NOT Output_A_Reset_TON[23].Q;
Out_CYw_Disc_Chk_A_H := _p126;
Output_A_M[23] := _p126;
(* Rung 101 *)
Out_CYw_Disc_Chk_A_H_Done := Output_A_M[23] AND TimerQ_In_SenCY_Disc_Chk_A_H;
Output_A_Reset_TON[23](In := Output_A_M[23] AND TimerQ_In_SenCY_Disc_Chk_A_H, PT := T#1s);
(* Rung 102 *)
Output_A_Error_TON[23](In := Out_CYw_Disc_Chk_A_H_Auto[1] AND AutoMode AND NOT Pause[1] AND NOT TimerQ_In_SenCY_Disc_Chk_A_H, PT := T#10s);
_e127(CLK := Output_A_Error_TON[23].Q);
IF _e127.Q THEN
    Output_A_Error_M[23] := TRUE;
    HMI_MessageNo[0] := INT#29;
END_IF;
(* Rung 103: 【Y717】排出A(左側)チャック開 行 *)
_e128(CLK := Out_CYw_Disc_Chk_A_F_Auto[1] AND AutoMode AND NOT Pause[1]);
_e129(CLK := Out_CYw_Disc_Chk_A_F_Manual[1] AND ManualMode);
_p130 := (_e128.Q OR _e129.Q OR Output_A_M[24]) AND NOT M9999 AND NOT Pause[1] AND NOT Output_A_Reset_TON[24].Q;
Out_CYw_Disc_Chk_A_F := _p130;
Output_A_M[24] := _p130;
(* Rung 104 *)
Out_CYw_Disc_Chk_A_F_Done := Output_A_M[24] AND TimerQ_In_SenCY_Disc_Chk_A_F;
Output_A_Reset_TON[24](In := Output_A_M[24] AND TimerQ_In_SenCY_Disc_Chk_A_F, PT := T#1s);

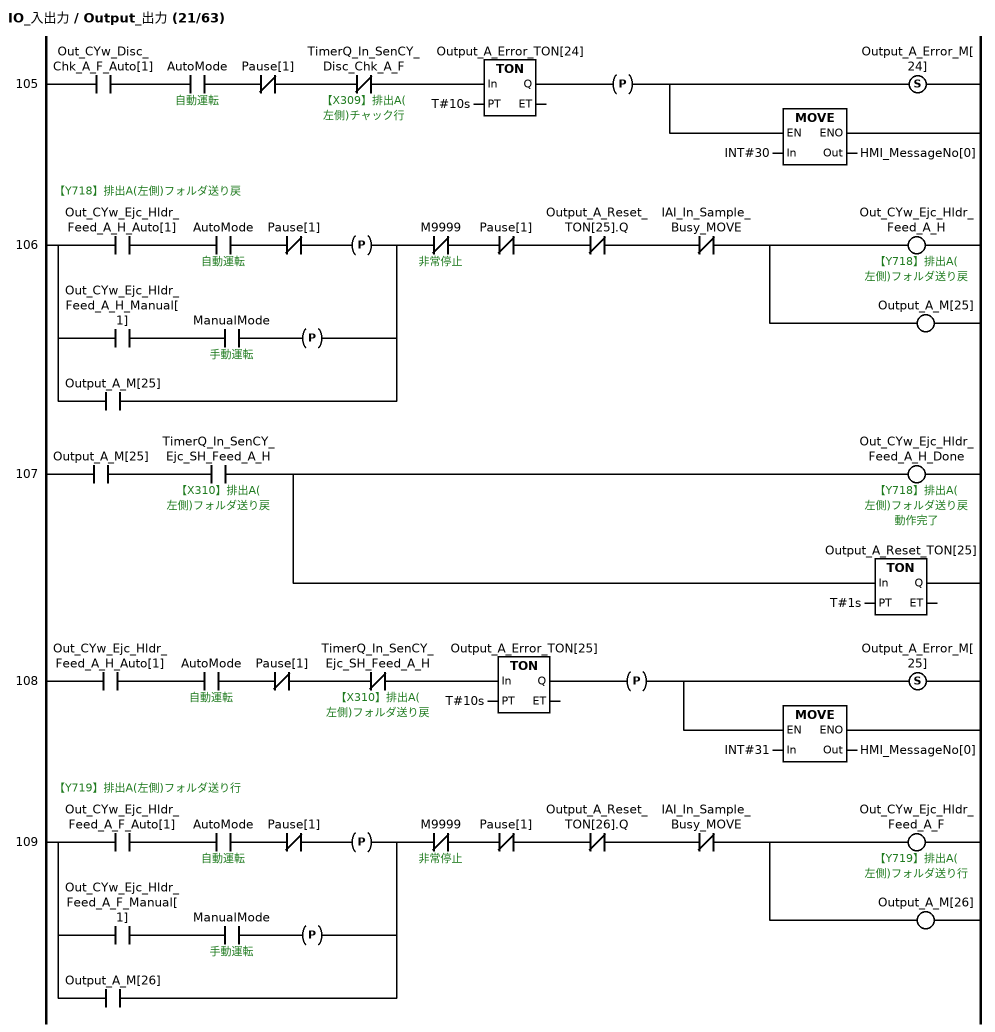
(* Rung 105 *)
Output_A_Error_TON[24](In := Out_CYw_Disc_Chk_A_F_Auto[1] AND AutoMode AND NOT Pause[1] AND NOT TimerQ_In_SenCY_Disc_Chk_A_F, PT := T#10s);
_e131(CLK := Output_A_Error_TON[24].Q);
IF _e131.Q THEN
    Output_A_Error_M[24] := TRUE;
    HMI_MessageNo[0] := INT#30;
END_IF;
(* Rung 106: 【Y718】排出A(左側)フォルダ送り戻 *)
_e132(CLK := Out_CYw_Ejc_Hldr_Feed_A_H_Auto[1] AND AutoMode AND NOT Pause[1]);
_e133(CLK := Out_CYw_Ejc_Hldr_Feed_A_H_Manual[1] AND ManualMode);
_p134 := (_e132.Q OR _e133.Q OR Output_A_M[25]) AND NOT M9999 AND NOT Pause[1] AND NOT Output_A_Reset_TON[25].Q AND NOT IAI_In_Sample_Busy_MOVE;
Out_CYw_Ejc_Hldr_Feed_A_H := _p134;
Output_A_M[25] := _p134;
(* Rung 107 *)
_p135 := Output_A_M[25] AND TimerQ_In_SenCY_Ejc_SH_Feed_A_H;
Out_CYw_Ejc_Hldr_Feed_A_H_Done := _p135;
Output_A_Reset_TON[25](In := _p135, PT := T#1s);
(* Rung 108 *)
Output_A_Error_TON[25](In := Out_CYw_Ejc_Hldr_Feed_A_H_Auto[1] AND AutoMode AND NOT Pause[1] AND NOT TimerQ_In_SenCY_Ejc_SH_Feed_A_H, PT := T#10s);
_e136(CLK := Output_A_Error_TON[25].Q);
IF _e136.Q THEN
    Output_A_Error_M[25] := TRUE;
    HMI_MessageNo[0] := INT#31;
END_IF;
(* Rung 109: 【Y719】排出A(左側)フォルダ送り行 *)
_e137(CLK := Out_CYw_Ejc_Hldr_Feed_A_F_Auto[1] AND AutoMode AND NOT Pause[1]);
_e138(CLK := Out_CYw_Ejc_Hldr_Feed_A_F_Manual[1] AND ManualMode);
_p139 := (_e137.Q OR _e138.Q OR Output_A_M[26]) AND NOT M9999 AND NOT Pause[1] AND NOT Output_A_Reset_TON[26].Q AND NOT IAI_In_Sample_Busy_MOVE;
Out_CYw_Ejc_Hldr_Feed_A_F := _p139;
Output_A_M[26] := _p139;

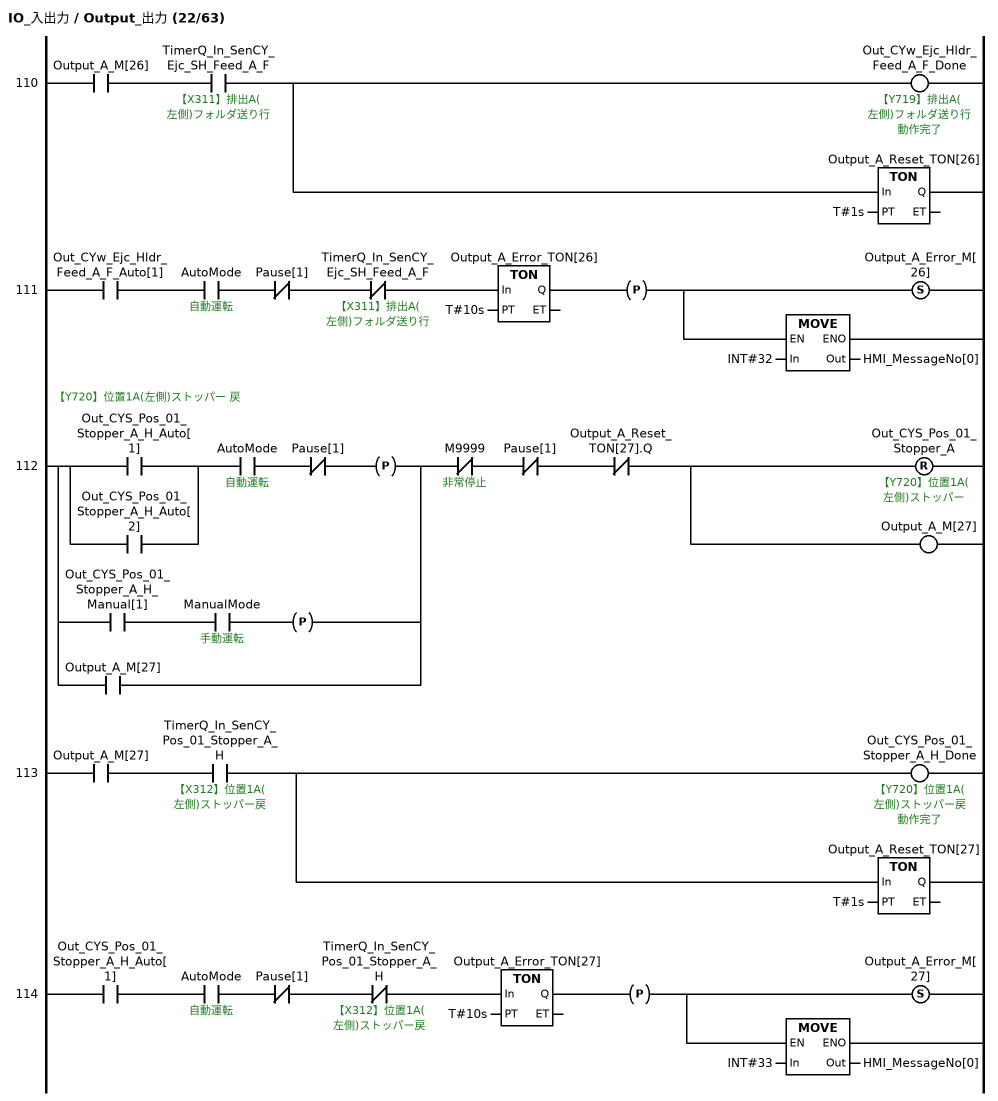
(* Rung 110 *)
_p140 := Output_A_M[26] AND TimerQ_In_SenCY_Ejc_SH_Feed_A_F;
Out_CYw_Ejc_Hldr_Feed_A_F_Done := _p140;
Output_A_Reset_TON[26](In := _p140, PT := T#1s);
(* Rung 111 *)
Output_A_Error_TON[26](In := Out_CYw_Ejc_Hldr_Feed_A_F_Auto[1] AND AutoMode AND NOT Pause[1] AND NOT TimerQ_In_SenCY_Ejc_SH_Feed_A_F, PT := T#10s);
_e141(CLK := Output_A_Error_TON[26].Q);
IF _e141.Q THEN
    Output_A_Error_M[26] := TRUE;
    HMI_MessageNo[0] := INT#32;
END_IF;
(* Rung 112: 【Y720】位置1A(左側)ストッパー 戻 *)
_e142(CLK := (Out_CYS_Pos_01_Stopper_A_H_Auto[1] OR Out_CYS_Pos_01_Stopper_A_H_Auto[2]) AND AutoMode AND NOT Pause[1]);
_e143(CLK := Out_CYS_Pos_01_Stopper_A_H_Manual[1] AND ManualMode);
_p144 := (_e142.Q OR _e143.Q OR Output_A_M[27]) AND NOT M9999 AND NOT Pause[1] AND NOT Output_A_Reset_TON[27].Q;
IF _p144 THEN Out_CYS_Pos_01_Stopper_A := FALSE; END_IF;
Output_A_M[27] := _p144;
(* Rung 113 *)
_p145 := Output_A_M[27] AND TimerQ_In_SenCY_Pos_01_Stopper_A_H;
Out_CYS_Pos_01_Stopper_A_H_Done := _p145;
Output_A_Reset_TON[27](In := _p145, PT := T#1s);
(* Rung 114 *)
Output_A_Error_TON[27](In := Out_CYS_Pos_01_Stopper_A_H_Auto[1] AND AutoMode AND NOT Pause[1] AND NOT TimerQ_In_SenCY_Pos_01_Stopper_A_H, PT := T#10s);
_e146(CLK := Output_A_Error_TON[27].Q);
IF _e146.Q THEN
    Output_A_Error_M[27] := TRUE;
    HMI_MessageNo[0] := INT#33;
END_IF;

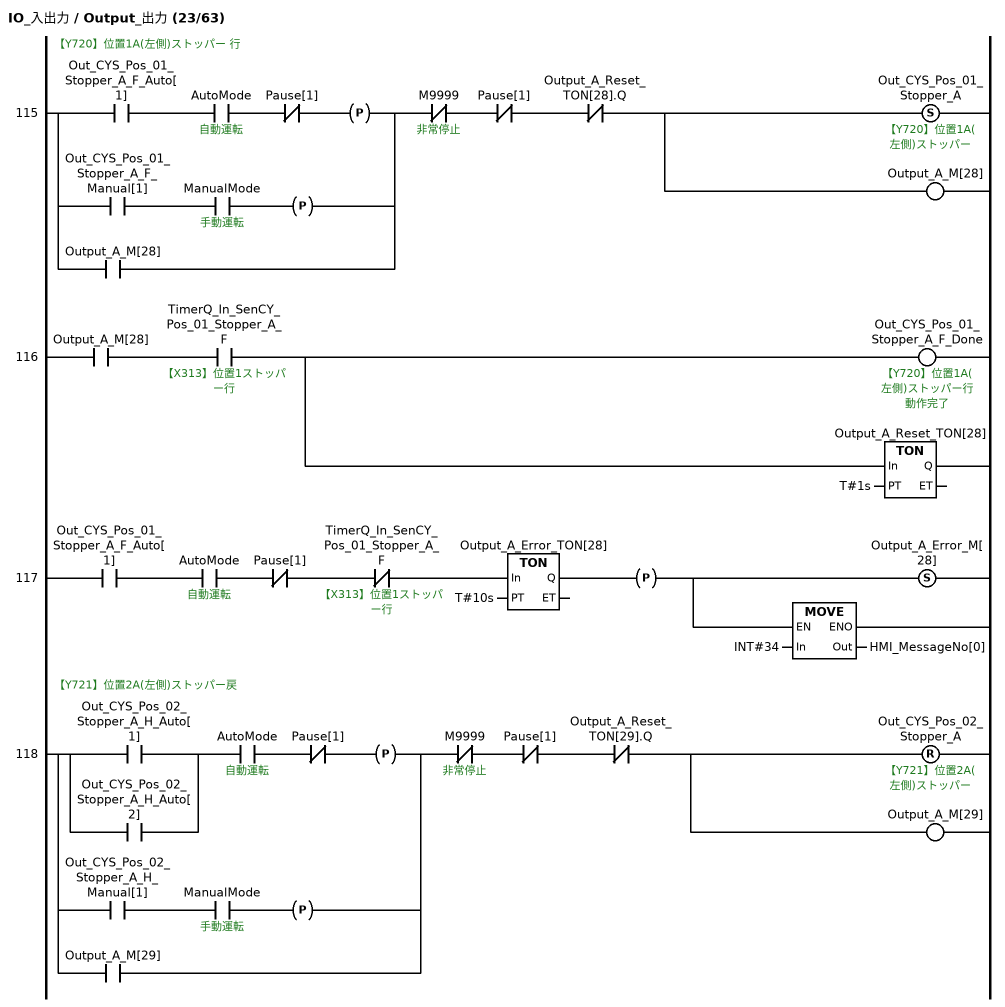
(* Rung 115: 【Y720】位置1A(左側)ストッパー 行 *)
_e147(CLK := Out_CYS_Pos_01_Stopper_A_F_Auto[1] AND AutoMode AND NOT Pause[1]);
_e148(CLK := Out_CYS_Pos_01_Stopper_A_F_Manual[1] AND ManualMode);
_p149 := (_e147.Q OR _e148.Q OR Output_A_M[28]) AND NOT M9999 AND NOT Pause[1] AND NOT Output_A_Reset_TON[28].Q;
IF _p149 THEN Out_CYS_Pos_01_Stopper_A := TRUE; END_IF;
Output_A_M[28] := _p149;
(* Rung 116 *)
_p150 := Output_A_M[28] AND TimerQ_In_SenCY_Pos_01_Stopper_A_F;
Out_CYS_Pos_01_Stopper_A_F_Done := _p150;
Output_A_Reset_TON[28](In := _p150, PT := T#1s);
(* Rung 117 *)
Output_A_Error_TON[28](In := Out_CYS_Pos_01_Stopper_A_F_Auto[1] AND AutoMode AND NOT Pause[1] AND NOT TimerQ_In_SenCY_Pos_01_Stopper_A_F, PT := T#10s);
_e151(CLK := Output_A_Error_TON[28].Q);
IF _e151.Q THEN
    Output_A_Error_M[28] := TRUE;
    HMI_MessageNo[0] := INT#34;
END_IF;
(* Rung 118: 【Y721】位置2A(左側)ストッパー戻 *)
_e152(CLK := (Out_CYS_Pos_02_Stopper_A_H_Auto[1] OR Out_CYS_Pos_02_Stopper_A_H_Auto[2]) AND AutoMode AND NOT Pause[1]);
_e153(CLK := Out_CYS_Pos_02_Stopper_A_H_Manual[1] AND ManualMode);
_p154 := (_e152.Q OR _e153.Q OR Output_A_M[29]) AND NOT M9999 AND NOT Pause[1] AND NOT Output_A_Reset_TON[29].Q;
IF _p154 THEN Out_CYS_Pos_02_Stopper_A := FALSE; END_IF;
Output_A_M[29] := _p154;

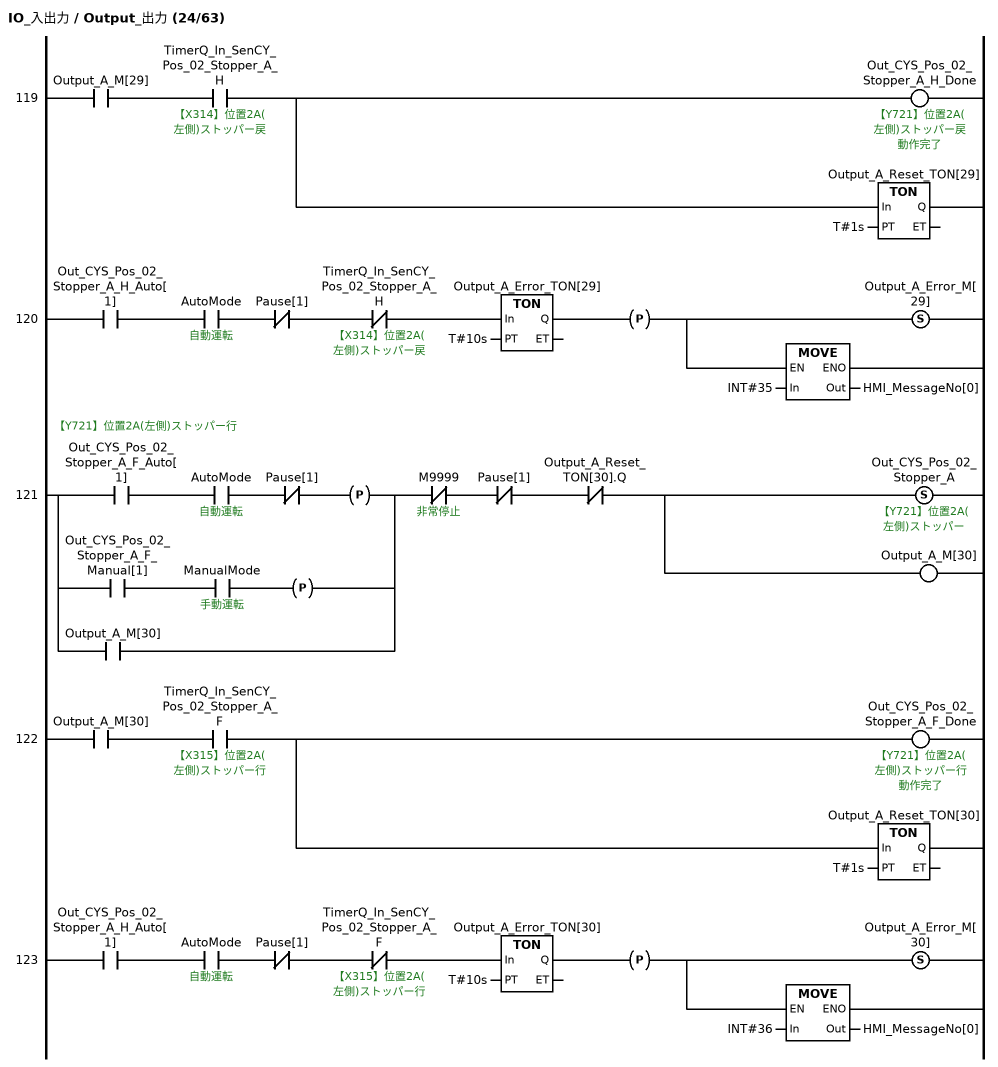
(* Rung 119 *)
_p155 := Output_A_M[29] AND TimerQ_In_SenCY_Pos_02_Stopper_A_H;
Out_CYS_Pos_02_Stopper_A_H_Done := _p155;
Output_A_Reset_TON[29](In := _p155, PT := T#1s);
(* Rung 120 *)
Output_A_Error_TON[29](In := Out_CYS_Pos_02_Stopper_A_H_Auto[1] AND AutoMode AND NOT Pause[1] AND NOT TimerQ_In_SenCY_Pos_02_Stopper_A_H, PT := T#10s);
_e156(CLK := Output_A_Error_TON[29].Q);
IF _e156.Q THEN
    Output_A_Error_M[29] := TRUE;
    HMI_MessageNo[0] := INT#35;
END_IF;
(* Rung 121: 【Y721】位置2A(左側)ストッパー行 *)
_e157(CLK := Out_CYS_Pos_02_Stopper_A_F_Auto[1] AND AutoMode AND NOT Pause[1]);
_e158(CLK := Out_CYS_Pos_02_Stopper_A_F_Manual[1] AND ManualMode);
_p159 := (_e157.Q OR _e158.Q OR Output_A_M[30]) AND NOT M9999 AND NOT Pause[1] AND NOT Output_A_Reset_TON[30].Q;
IF _p159 THEN Out_CYS_Pos_02_Stopper_A := TRUE; END_IF;
Output_A_M[30] := _p159;
(* Rung 122 *)
_p160 := Output_A_M[30] AND TimerQ_In_SenCY_Pos_02_Stopper_A_F;
Out_CYS_Pos_02_Stopper_A_F_Done := _p160;
Output_A_Reset_TON[30](In := _p160, PT := T#1s);
(* Rung 123 *)
Output_A_Error_TON[30](In := Out_CYS_Pos_02_Stopper_A_H_Auto[1] AND AutoMode AND NOT Pause[1] AND NOT TimerQ_In_SenCY_Pos_02_Stopper_A_F, PT := T#10s);
_e161(CLK := Output_A_Error_TON[30].Q);
IF _e161.Q THEN
    Output_A_Error_M[30] := TRUE;
    HMI_MessageNo[0] := INT#36;
END_IF;

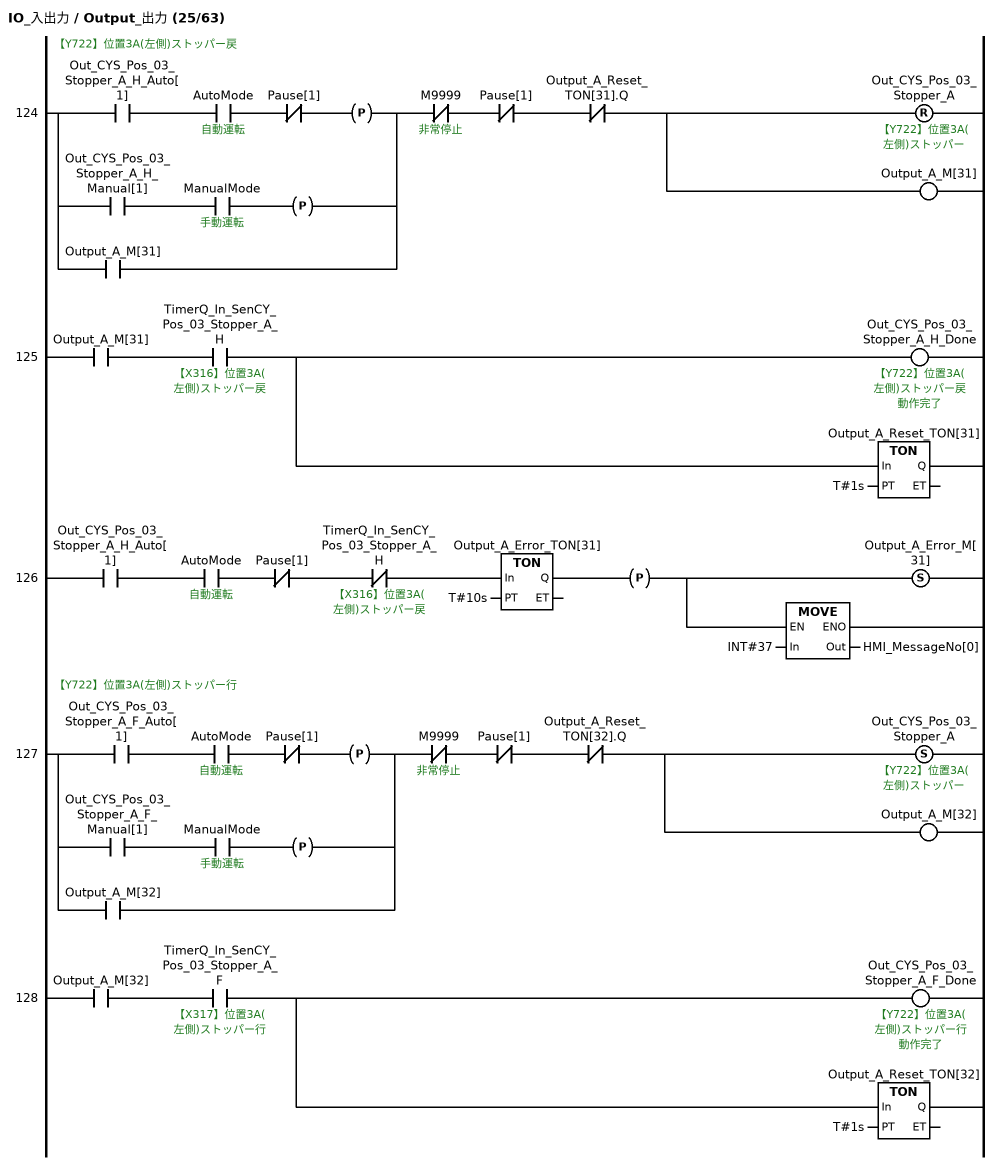
(* Rung 124: 【Y722】位置3A(左側)ストッパー戻 *)
_e162(CLK := Out_CYS_Pos_03_Stopper_A_H_Auto[1] AND AutoMode AND NOT Pause[1]);
_e163(CLK := Out_CYS_Pos_03_Stopper_A_H_Manual[1] AND ManualMode);
_p164 := (_e162.Q OR _e163.Q OR Output_A_M[31]) AND NOT M9999 AND NOT Pause[1] AND NOT Output_A_Reset_TON[31].Q;
IF _p164 THEN Out_CYS_Pos_03_Stopper_A := FALSE; END_IF;
Output_A_M[31] := _p164;
(* Rung 125 *)
_p165 := Output_A_M[31] AND TimerQ_In_SenCY_Pos_03_Stopper_A_H;
Out_CYS_Pos_03_Stopper_A_H_Done := _p165;
Output_A_Reset_TON[31](In := _p165, PT := T#1s);
(* Rung 126 *)
Output_A_Error_TON[31](In := Out_CYS_Pos_03_Stopper_A_H_Auto[1] AND AutoMode AND NOT Pause[1] AND NOT TimerQ_In_SenCY_Pos_03_Stopper_A_H, PT := T#10s);
_e166(CLK := Output_A_Error_TON[31].Q);
IF _e166.Q THEN
    Output_A_Error_M[31] := TRUE;
    HMI_MessageNo[0] := INT#37;
END_IF;
(* Rung 127: 【Y722】位置3A(左側)ストッパー行 *)
_e167(CLK := Out_CYS_Pos_03_Stopper_A_F_Auto[1] AND AutoMode AND NOT Pause[1]);
_e168(CLK := Out_CYS_Pos_03_Stopper_A_F_Manual[1] AND ManualMode);
_p169 := (_e167.Q OR _e168.Q OR Output_A_M[32]) AND NOT M9999 AND NOT Pause[1] AND NOT Output_A_Reset_TON[32].Q;
IF _p169 THEN Out_CYS_Pos_03_Stopper_A := TRUE; END_IF;
Output_A_M[32] := _p169;
(* Rung 128 *)
_p170 := Output_A_M[32] AND TimerQ_In_SenCY_Pos_03_Stopper_A_F;
Out_CYS_Pos_03_Stopper_A_F_Done := _p170;
Output_A_Reset_TON[32](In := _p170, PT := T#1s);

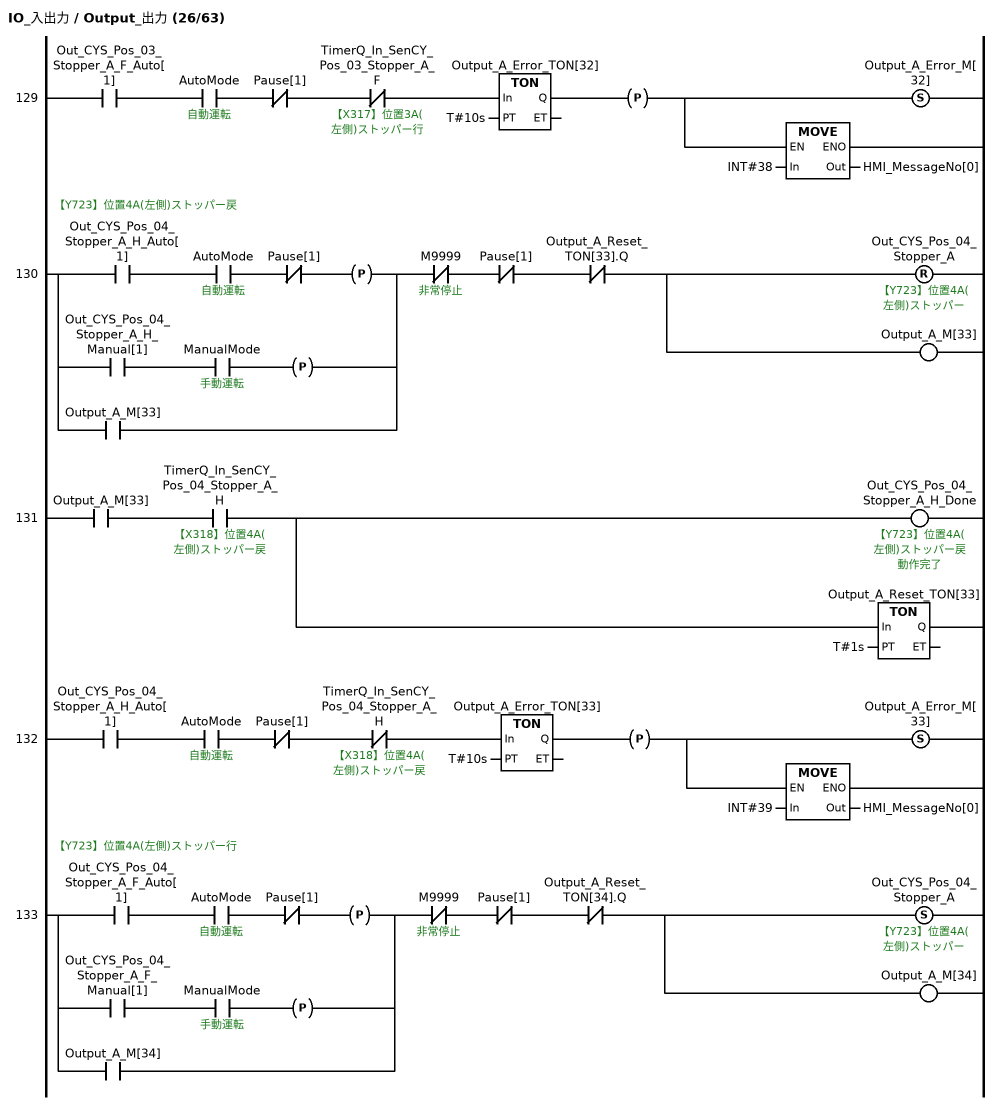
(* Rung 129 *)
Output_A_Error_TON[32](In := Out_CYS_Pos_03_Stopper_A_F_Auto[1] AND AutoMode AND NOT Pause[1] AND NOT TimerQ_In_SenCY_Pos_03_Stopper_A_F, PT := T#10s);
_e171(CLK := Output_A_Error_TON[32].Q);
IF _e171.Q THEN
    Output_A_Error_M[32] := TRUE;
    HMI_MessageNo[0] := INT#38;
END_IF;
(* Rung 130: 【Y723】位置4A(左側)ストッパー戻 *)
_e172(CLK := Out_CYS_Pos_04_Stopper_A_H_Auto[1] AND AutoMode AND NOT Pause[1]);
_e173(CLK := Out_CYS_Pos_04_Stopper_A_H_Manual[1] AND ManualMode);
_p174 := (_e172.Q OR _e173.Q OR Output_A_M[33]) AND NOT M9999 AND NOT Pause[1] AND NOT Output_A_Reset_TON[33].Q;
IF _p174 THEN Out_CYS_Pos_04_Stopper_A := FALSE; END_IF;
Output_A_M[33] := _p174;
(* Rung 131 *)
_p175 := Output_A_M[33] AND TimerQ_In_SenCY_Pos_04_Stopper_A_H;
Out_CYS_Pos_04_Stopper_A_H_Done := _p175;
Output_A_Reset_TON[33](In := _p175, PT := T#1s);
(* Rung 132 *)
Output_A_Error_TON[33](In := Out_CYS_Pos_04_Stopper_A_H_Auto[1] AND AutoMode AND NOT Pause[1] AND NOT TimerQ_In_SenCY_Pos_04_Stopper_A_H, PT := T#10s);
_e176(CLK := Output_A_Error_TON[33].Q);
IF _e176.Q THEN
    Output_A_Error_M[33] := TRUE;
    HMI_MessageNo[0] := INT#39;
END_IF;
(* Rung 133: 【Y723】位置4A(左側)ストッパー行 *)
_e177(CLK := Out_CYS_Pos_04_Stopper_A_F_Auto[1] AND AutoMode AND NOT Pause[1]);
_e178(CLK := Out_CYS_Pos_04_Stopper_A_F_Manual[1] AND ManualMode);
_p179 := (_e177.Q OR _e178.Q OR Output_A_M[34]) AND NOT M9999 AND NOT Pause[1] AND NOT Output_A_Reset_TON[34].Q;
IF _p179 THEN Out_CYS_Pos_04_Stopper_A := TRUE; END_IF;
Output_A_M[34] := _p179;

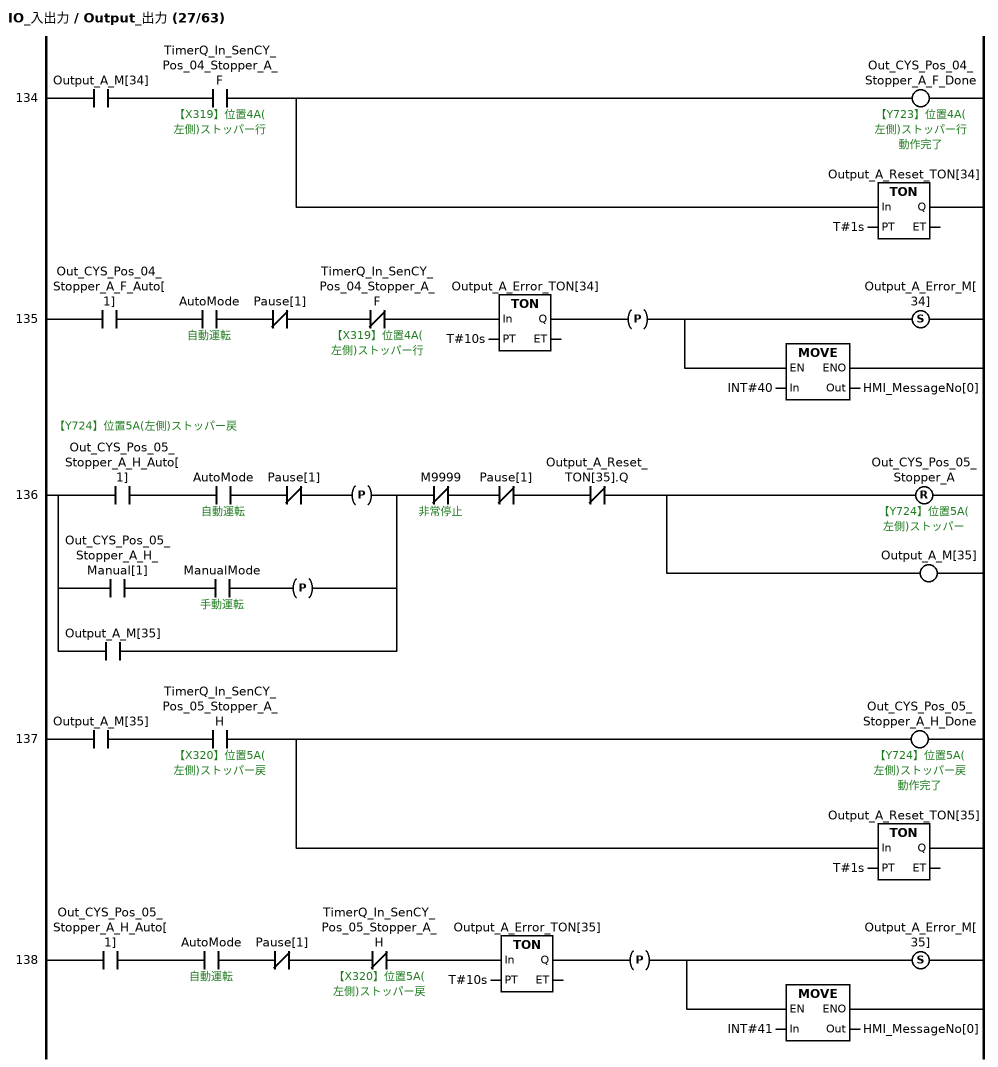
(* Rung 134 *)
_p180 := Output_A_M[34] AND TimerQ_In_SenCY_Pos_04_Stopper_A_F;
Out_CYS_Pos_04_Stopper_A_F_Done := _p180;
Output_A_Reset_TON[34](In := _p180, PT := T#1s);
(* Rung 135 *)
Output_A_Error_TON[34](In := Out_CYS_Pos_04_Stopper_A_F_Auto[1] AND AutoMode AND NOT Pause[1] AND NOT TimerQ_In_SenCY_Pos_04_Stopper_A_F, PT := T#10s);
_e181(CLK := Output_A_Error_TON[34].Q);
IF _e181.Q THEN
    Output_A_Error_M[34] := TRUE;
    HMI_MessageNo[0] := INT#40;
END_IF;
(* Rung 136: 【Y724】位置5A(左側)ストッパー戻 *)
_e182(CLK := Out_CYS_Pos_05_Stopper_A_H_Auto[1] AND AutoMode AND NOT Pause[1]);
_e183(CLK := Out_CYS_Pos_05_Stopper_A_H_Manual[1] AND ManualMode);
_p184 := (_e182.Q OR _e183.Q OR Output_A_M[35]) AND NOT M9999 AND NOT Pause[1] AND NOT Output_A_Reset_TON[35].Q;
IF _p184 THEN Out_CYS_Pos_05_Stopper_A := FALSE; END_IF;
Output_A_M[35] := _p184;
(* Rung 137 *)
_p185 := Output_A_M[35] AND TimerQ_In_SenCY_Pos_05_Stopper_A_H;
Out_CYS_Pos_05_Stopper_A_H_Done := _p185;
Output_A_Reset_TON[35](In := _p185, PT := T#1s);
(* Rung 138 *)
Output_A_Error_TON[35](In := Out_CYS_Pos_05_Stopper_A_H_Auto[1] AND AutoMode AND NOT Pause[1] AND NOT TimerQ_In_SenCY_Pos_05_Stopper_A_H, PT := T#10s);
_e186(CLK := Output_A_Error_TON[35].Q);
IF _e186.Q THEN
    Output_A_Error_M[35] := TRUE;
    HMI_MessageNo[0] := INT#41;
END_IF;

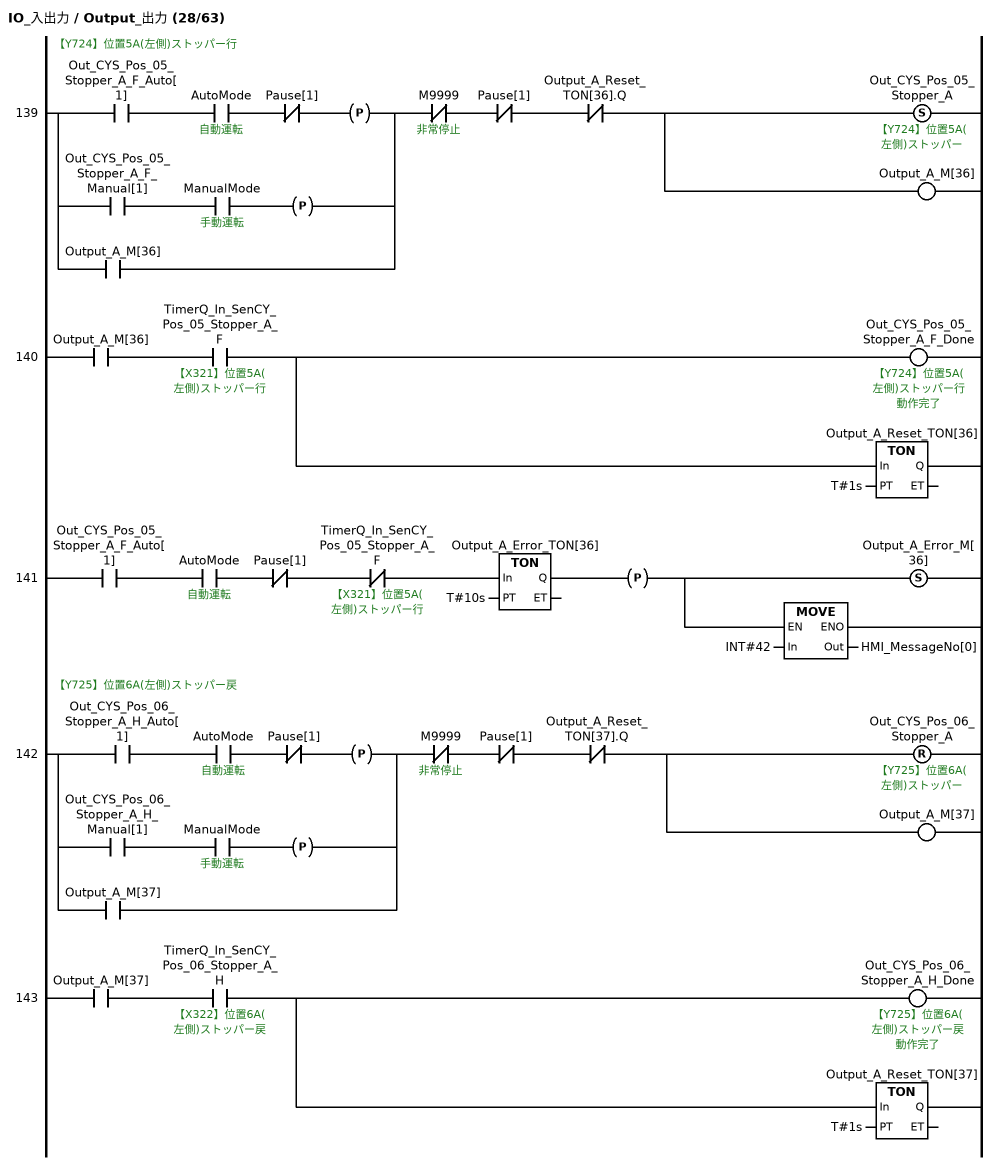
(* Rung 139: 【Y724】位置5A(左側)ストッパー行 *)
_e187(CLK := Out_CYS_Pos_05_Stopper_A_F_Auto[1] AND AutoMode AND NOT Pause[1]);
_e188(CLK := Out_CYS_Pos_05_Stopper_A_F_Manual[1] AND ManualMode);
_p189 := (_e187.Q OR _e188.Q OR Output_A_M[36]) AND NOT M9999 AND NOT Pause[1] AND NOT Output_A_Reset_TON[36].Q;
IF _p189 THEN Out_CYS_Pos_05_Stopper_A := TRUE; END_IF;
Output_A_M[36] := _p189;
(* Rung 140 *)
_p190 := Output_A_M[36] AND TimerQ_In_SenCY_Pos_05_Stopper_A_F;
Out_CYS_Pos_05_Stopper_A_F_Done := _p190;
Output_A_Reset_TON[36](In := _p190, PT := T#1s);
(* Rung 141 *)
Output_A_Error_TON[36](In := Out_CYS_Pos_05_Stopper_A_F_Auto[1] AND AutoMode AND NOT Pause[1] AND NOT TimerQ_In_SenCY_Pos_05_Stopper_A_F, PT := T#10s);
_e191(CLK := Output_A_Error_TON[36].Q);
IF _e191.Q THEN
    Output_A_Error_M[36] := TRUE;
    HMI_MessageNo[0] := INT#42;
END_IF;
(* Rung 142: 【Y725】位置6A(左側)ストッパー戻 *)
_e192(CLK := Out_CYS_Pos_06_Stopper_A_H_Auto[1] AND AutoMode AND NOT Pause[1]);
_e193(CLK := Out_CYS_Pos_06_Stopper_A_H_Manual[1] AND ManualMode);
_p194 := (_e192.Q OR _e193.Q OR Output_A_M[37]) AND NOT M9999 AND NOT Pause[1] AND NOT Output_A_Reset_TON[37].Q;
IF _p194 THEN Out_CYS_Pos_06_Stopper_A := FALSE; END_IF;
Output_A_M[37] := _p194;
(* Rung 143 *)
_p195 := Output_A_M[37] AND TimerQ_In_SenCY_Pos_06_Stopper_A_H;
Out_CYS_Pos_06_Stopper_A_H_Done := _p195;
Output_A_Reset_TON[37](In := _p195, PT := T#1s);

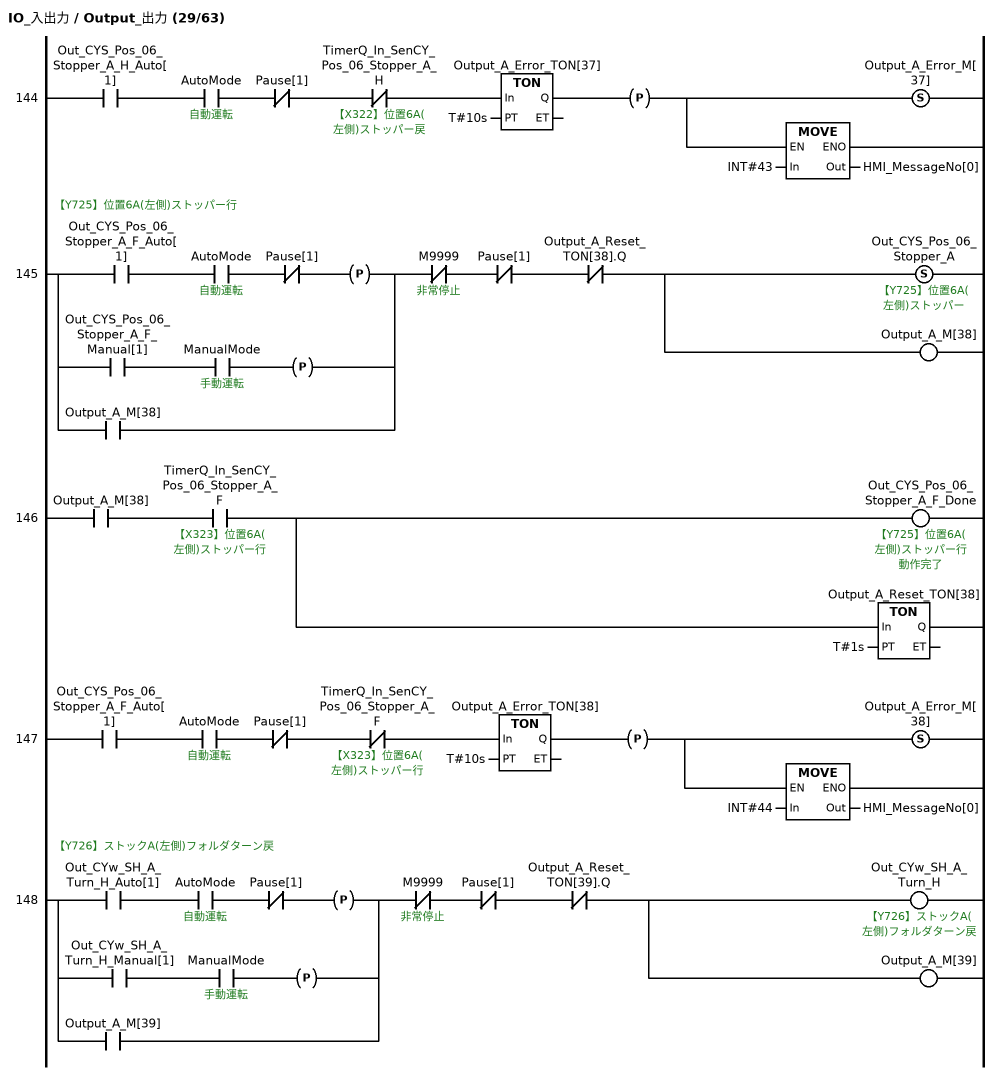
(* Rung 144 *)
Output_A_Error_TON[37](In := Out_CYS_Pos_06_Stopper_A_H_Auto[1] AND AutoMode AND NOT Pause[1] AND NOT TimerQ_In_SenCY_Pos_06_Stopper_A_H, PT := T#10s);
_e196(CLK := Output_A_Error_TON[37].Q);
IF _e196.Q THEN
    Output_A_Error_M[37] := TRUE;
    HMI_MessageNo[0] := INT#43;
END_IF;
(* Rung 145: 【Y725】位置6A(左側)ストッパー行 *)
_e197(CLK := Out_CYS_Pos_06_Stopper_A_F_Auto[1] AND AutoMode AND NOT Pause[1]);
_e198(CLK := Out_CYS_Pos_06_Stopper_A_F_Manual[1] AND ManualMode);
_p199 := (_e197.Q OR _e198.Q OR Output_A_M[38]) AND NOT M9999 AND NOT Pause[1] AND NOT Output_A_Reset_TON[38].Q;
IF _p199 THEN Out_CYS_Pos_06_Stopper_A := TRUE; END_IF;
Output_A_M[38] := _p199;
(* Rung 146 *)
_p200 := Output_A_M[38] AND TimerQ_In_SenCY_Pos_06_Stopper_A_F;
Out_CYS_Pos_06_Stopper_A_F_Done := _p200;
Output_A_Reset_TON[38](In := _p200, PT := T#1s);
(* Rung 147 *)
Output_A_Error_TON[38](In := Out_CYS_Pos_06_Stopper_A_F_Auto[1] AND AutoMode AND NOT Pause[1] AND NOT TimerQ_In_SenCY_Pos_06_Stopper_A_F, PT := T#10s);
_e201(CLK := Output_A_Error_TON[38].Q);
IF _e201.Q THEN
    Output_A_Error_M[38] := TRUE;
    HMI_MessageNo[0] := INT#44;
END_IF;
(* Rung 148: 【Y726】ストックA(左側)フォルダターン戻 *)
_e202(CLK := Out_CYw_SH_A_Turn_H_Auto[1] AND AutoMode AND NOT Pause[1]);
_e203(CLK := Out_CYw_SH_A_Turn_H_Manual[1] AND ManualMode);
_p204 := (_e202.Q OR _e203.Q OR Output_A_M[39]) AND NOT M9999 AND NOT Pause[1] AND NOT Output_A_Reset_TON[39].Q;
Out_CYw_SH_A_Turn_H := _p204;
Output_A_M[39] := _p204;

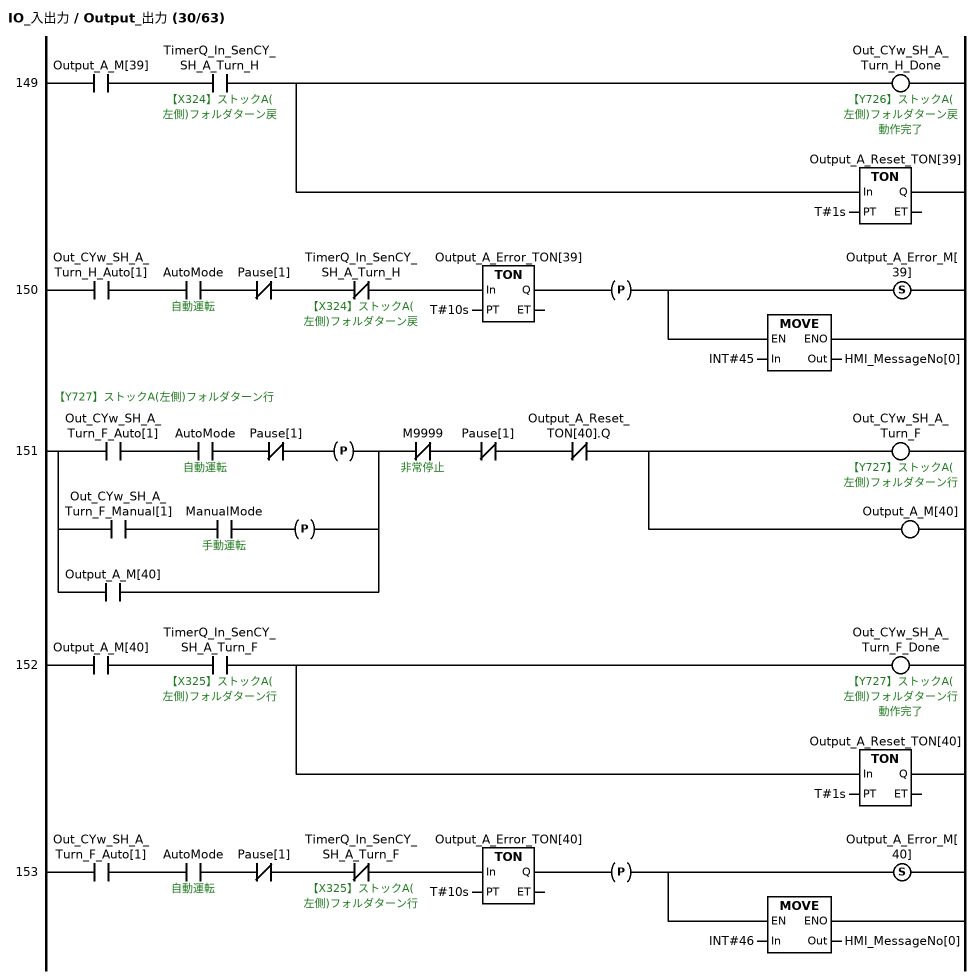
(* Rung 149 *)
Out_CYw_SH_A_Turn_H_Done := Output_A_M[39] AND TimerQ_In_SenCY_SH_A_Turn_H;
Output_A_Reset_TON[39](In := Output_A_M[39] AND TimerQ_In_SenCY_SH_A_Turn_H, PT := T#1s);
(* Rung 150 *)
Output_A_Error_TON[39](In := Out_CYw_SH_A_Turn_H_Auto[1] AND AutoMode AND NOT Pause[1] AND NOT TimerQ_In_SenCY_SH_A_Turn_H, PT := T#10s);
_e205(CLK := Output_A_Error_TON[39].Q);
IF _e205.Q THEN
    Output_A_Error_M[39] := TRUE;
    HMI_MessageNo[0] := INT#45;
END_IF;
(* Rung 151: 【Y727】ストックA(左側)フォルダターン行 *)
_e206(CLK := Out_CYw_SH_A_Turn_F_Auto[1] AND AutoMode AND NOT Pause[1]);
_e207(CLK := Out_CYw_SH_A_Turn_F_Manual[1] AND ManualMode);
_p208 := (_e206.Q OR _e207.Q OR Output_A_M[40]) AND NOT M9999 AND NOT Pause[1] AND NOT Output_A_Reset_TON[40].Q;
Out_CYw_SH_A_Turn_F := _p208;
Output_A_M[40] := _p208;
(* Rung 152 *)
Out_CYw_SH_A_Turn_F_Done := Output_A_M[40] AND TimerQ_In_SenCY_SH_A_Turn_F;
Output_A_Reset_TON[40](In := Output_A_M[40] AND TimerQ_In_SenCY_SH_A_Turn_F, PT := T#1s);
(* Rung 153 *)
Output_A_Error_TON[40](In := Out_CYw_SH_A_Turn_F_Auto[1] AND AutoMode AND NOT Pause[1] AND NOT TimerQ_In_SenCY_SH_A_Turn_F, PT := T#10s);
_e209(CLK := Output_A_Error_TON[40].Q);
IF _e209.Q THEN
    Output_A_Error_M[40] := TRUE;
    HMI_MessageNo[0] := INT#46;
END_IF;

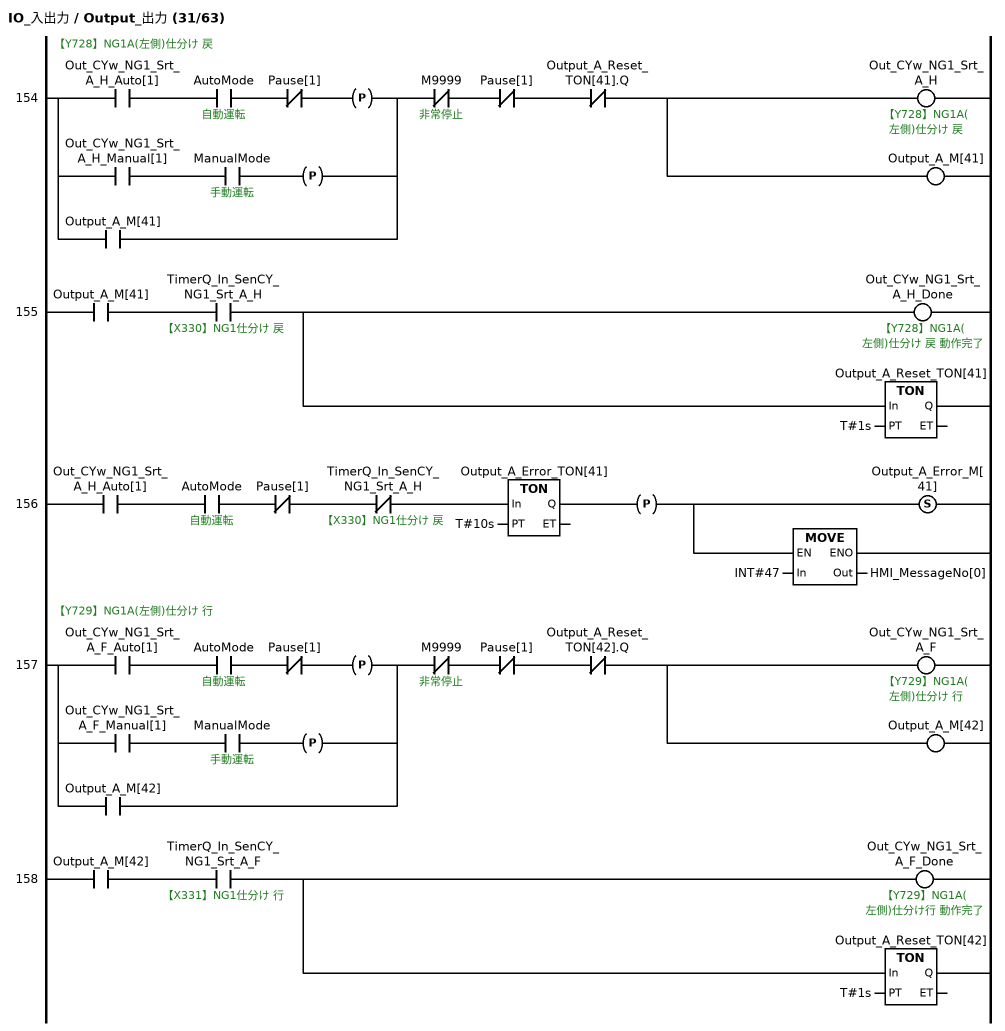
(* Rung 154: 【Y728】NG1A(左側)仕分け 戻 *)
_e210(CLK := Out_CYw_NG1_Srt_A_H_Auto[1] AND AutoMode AND NOT Pause[1]);
_e211(CLK := Out_CYw_NG1_Srt_A_H_Manual[1] AND ManualMode);
_p212 := (_e210.Q OR _e211.Q OR Output_A_M[41]) AND NOT M9999 AND NOT Pause[1] AND NOT Output_A_Reset_TON[41].Q;
Out_CYw_NG1_Srt_A_H := _p212;
Output_A_M[41] := _p212;
(* Rung 155 *)
Out_CYw_NG1_Srt_A_H_Done := Output_A_M[41] AND TimerQ_In_SenCY_NG1_Srt_A_H;
Output_A_Reset_TON[41](In := Output_A_M[41] AND TimerQ_In_SenCY_NG1_Srt_A_H, PT := T#1s);
(* Rung 156 *)
Output_A_Error_TON[41](In := Out_CYw_NG1_Srt_A_H_Auto[1] AND AutoMode AND NOT Pause[1] AND NOT TimerQ_In_SenCY_NG1_Srt_A_H, PT := T#10s);
_e213(CLK := Output_A_Error_TON[41].Q);
IF _e213.Q THEN
    Output_A_Error_M[41] := TRUE;
    HMI_MessageNo[0] := INT#47;
END_IF;
(* Rung 157: 【Y729】NG1A(左側)仕分け 行 *)
_e214(CLK := Out_CYw_NG1_Srt_A_F_Auto[1] AND AutoMode AND NOT Pause[1]);
_e215(CLK := Out_CYw_NG1_Srt_A_F_Manual[1] AND ManualMode);
_p216 := (_e214.Q OR _e215.Q OR Output_A_M[42]) AND NOT M9999 AND NOT Pause[1] AND NOT Output_A_Reset_TON[42].Q;
Out_CYw_NG1_Srt_A_F := _p216;
Output_A_M[42] := _p216;
(* Rung 158 *)
Out_CYw_NG1_Srt_A_F_Done := Output_A_M[42] AND TimerQ_In_SenCY_NG1_Srt_A_F;
Output_A_Reset_TON[42](In := Output_A_M[42] AND TimerQ_In_SenCY_NG1_Srt_A_F, PT := T#1s);

